CASE nCode OF
	16#000 : sText := '0: No error  ';
	16#001 : sText := '1: Internal error  ';
	16#002 : sText := '2: No Rtime  ';
	16#003 : sText := '3: Allocation locked memory error  ';
	16#004 : sText := '4: Insert mailbox error  ';
	16#005 : sText := '5: Wrong receive HMSG  ';
	16#006 : sText := '6: target port not found  ';
	16#007 : sText := '7: target machine not found  ';
	16#008 : sText := '8: Unknown command ID  ';
	16#009 : sText := '9: Bad task ID  ';
	16#00A : sText := '10: No IO  ';
	16#00B : sText := '11: Unknown AMS command  ';
	16#00C : sText := '12: Win 32 error  ';
	16#00D : sText := '13: Port not connected  ';
	16#00E : sText := '14: Invalid AMS length  ';
	16#00F : sText := '15: Invalid AMS Net ID  ';
	16#010 : sText := '16: Low Installation level  ';
	16#011 : sText := '17: No debug available  ';
	16#012 : sText := '18: Port disabled  ';
	16#013 : sText := '19: Port already connected  ';
	16#014 : sText := '20: AMS Sync Win32 error  ';
	16#015 : sText := '21: AMS Sync Timeout  ';
	16#016 : sText := '22: AMS Sync AMS error  ';
	16#017 : sText := '23: AMS Sync no index map  '; 
	16#018 : sText := '24: Invalid AMS port  ';
	16#019 : sText := '25: No memory  ';
	16#01A : sText := '26: TCP send error  ';
	16#01B : sText := '27: Host unreachable  ';
	16#1000 : sText := '4096: Intern: RTERR_INTERNAL : $R$N Internal fatal error in the TwinCAT real-time system.  ';
	16#1001 : sText := '4097: Intern: RTERR_BADTIMERPERIODS: $R$N Timer value not vaild.  ';
	16#1002 : sText := '4098: Intern: RTERR_INVALIDTASKPTR: $R$N Task pointer has the invalid value ZERO. ';
	16#1003 : sText := '4099: Intern: RTERR_INVALIDSTACKPTR: $R$N Task stack pointer has the invalid value ZERO. ';
	16#1004 : sText := '4100: Intern: RTERR_PRIOEXISTS: $R$N The demand task priority is already assigned.  ';
	16#1005 : sText := '4101: Intern: RTERR_NOMORETCB: $R$N No more free TCB (Task Control Block) available. Maximum number of TCBs is 64.  ';
	16#1006 : sText := '4102: Intern: RTERR_NOMORESEMAS: $R$N No more free semaphores available. Maximum number of semaphores is 64.  ';
	16#1007 : sText := '4103: Intern: RTERR_NOMOREQUEUES: $R$N No more free queue available. Maximum number of queue is 64.  ';
	16#1008 : sText := '4104: Intern: TwinCAT reserved.:  ';
	16#1009 : sText := '4105: Intern: TwinCAT reserved.:  '; 
	16#100a : sText := '4106: Intern: TwinCAT reserved.:  '; 
	16#100b : sText := '4107: Intern: TwinCAT reserved.:  '; 
	16#100C : sText := '4108: Intern: TwinCAT reserved.:  ';
	16#100D : sText := '4109: Intern: RTERR_EXTIRQALREADYDEF: $R$N An external synchronisation interrupt is already applied. ';
	16#100E : sText := '4110: Intern: RTERR_EXTIRQNOTDEF: $R$N No external synchronsiation interrupt applied. ';
	16#100F : sText := '4111: Intern: RTERR_EXTIRQINSTALLFAILED: $R$N The apply of the external synchronisation interrupt failed. ';
	16#1010 : sText := '4112: Intern: RTERR_IRQLNOTLESSOREQUAL: $R$N Call of a service function in the wrong context.  ';
	16#2000 : sText := ': ERR_IOERRS  ';
	16#274C : sText := '10060: A socket operation was attempted to an unreachable host  ';
	16#274D : sText := '10061: A connection attempt failed because the connected party did not properly respond after a period of time, $R$N or established connection failed because connected host has failed to respond.  ';
	16#2751 : sText := '10065: No connection could be made because the target machine actively refused it  ';
	16#2900 : sText := ': ERR_DPSLAVE (ERR_IOERRS+0x900)  ';
	16#2A00 : sText := ': ERR_CP5412A2 (ERR_IOERRS+0xA00)  '; 
	16#2B00 : sText := ': ERR_ASP (ERR_IOERRS+0xB00)  '; 
	16#2C00 : sText := ': ERR_CANSLAVE (ERR_IOERRS+0xC00)  '; 
	16#2D00 : sText := ': ERR_CIF30 (ERR_IOERRS+0xD00)  '; 
	16#2E00 : sText := ': ERR_IBSSLAVE (ERR_IOERRS+0xE00)  ';
	16#3000 : sText := ': ERR_SPSERRS  '; 
	16#4000 : sText := ': ERR_NCERRS  ';
	16#500 : sText := '1280: Intern: ROUTERERR_NOLOCKEDMEMORY: $R$N No locked memory can be allocated.  ';
	16#501 : sText := '1281: Intern: ROUTERERR_RESIZEMEMORY: $R$N The size of the  router memory could not be changed. ';
	16#502 : sText := '1282: Intern: ROUTERERR_MAILBOXFULL: $R$N The Mailbox of the AmsPort has reached the maximum number of possible entries. The current sent message was abolished.  ';
	16#503 : sText := '1283: Intern: ROUTERERR_DEBUGBOXFULL: $R$N The Mailbox of the Ams debugger port has reached the maximum number of possible entries. $R$N The sent message wil not be displayed in the debug monitor.  ';
	16#504 : sText := '1284: Intern: ROUTERERR_UNKNOWNPORTTYPE :  ';
	16#505 : sText := '1285: Intern: ROUTERERR_NOTINITIALIZED: $R$N Router is not (yet) initialised.  ';
	16#506 : sText := '1286: Intern: ROUTERERR_PORTALREADYINUSE : $R$N The desired port number is already assigned. ';
	16#507 : sText := '1287: Intern: ROUTERERR_NOTREGISTERED : $R$N Ams Port not registered  ';
	16#508 : sText := '1288: Intern: ROUTERERR_NOMOREQUEUES: $R$N The maximum number of Ams Ports reached.  ';
	16#509 : sText := '1289: Intern: ROUTERERR_INVALIDPORT :  '; 
	16#50A : sText := '1290: Intern: ROUTERERR_NOTACTIVATED : $R$N TwinCAT Router not (yet) active.  ';
	16#6000 : sText := ': ERR_PLCERRS  ';
	16#0700 : sText := '1792: error class <device error>  ';
	16#7000 : sText := ': ERR_STRKERRS  '; 
	16#0701 : sText := '1793: Service is not supported by server  ';
	16#0702 : sText := '1794: invalid index group  ';
	16#0703 : sText := '1795: invalid index offset  ';
	16#0704 : sText := '1796: reading/writing not permitted  ';
	16#0705 : sText := '1797 : parameter size not correct  ';
	16#0706 : sText := '1798: invalid parameter value(s)  ';
	16#0707 : sText := '1799: device is not in a ready state  ';
	16#708 : sText := '1800: device is busy  '; 
	16#709 : sText := '1801: invalid context (must be in Windows)  ';
	16#70A : sText := '1802: out of memory  '; 
	16#70B : sText := '1803: invalid parameter value(s)  '; 
	16#70C : sText := '1804: not found (files, ...)  ';
	16#70D : sText := '1805: syntax error in command or file  '; 
	16#70E : sText := '1806: objects do not match  '; 
	16#70F : sText := '1807: object already exists  '; 
	16#710 : sText := '1808: symbol not found  '; 
	16#711 : sText := '1809: symbol version invalid  '; 
	16#712 : sText := '1810: server is in invalid state  '; 
	16#713 : sText := '1811: AdsTransMode not supported  '; 
	16#714 : sText := '1812: Notification handle is invalid  '; 
	16#715 : sText := '1813: Notification client not registered  '; 
	16#716 : sText := '1814: no more notification handles  '; 
	16#717 : sText := '1815: size for watch too big  ';
	16#718 : sText := '1816: device not initialized  ';
	16#719 : sText := '1817: device has a timeout  '; 
	16#71A : sText := '1818: query interface failed  '; 
	16#71B : sText := '1819: wrong interface required  '; 
	16#71C : sText := '1820: class ID is invalid  '; 
	16#71D : sText := '1821: object ID is invalid  '; 
	16#71E : sText := '1822: request is pending  '; 
	16#71F : sText := '1823: request is aborted  '; 
	16#720 : sText := '1824: signal warning  '; 
	16#721 : sText := '1825: invalid array index  ';
	16#722 : sText := '1826: symbol not active -> release handle and try again  ';
	16#723 : sText := '1827: access denied  ';
	16#740 : sText := '1856: Error class <client error>  ';
	16#741 : sText := '1857: invalid parameter at service  ';
	16#742 : sText := '1858: polling list is empty  '; 
	16#743 : sText := '1859: var connection already in use  ';
	16#744 : sText := '1860: invoke ID in use  ';
	16#745 : sText := '1861: timeout elapsed  ';
	16#746 : sText := '1862: error in win32 subsystem  '; 
	16#748 : sText := '1864: ads port not opened  '; 
	16#750 : sText := '1872: internal error in ads sync  ';
	16#751 : sText := '1873: hash table overflow  ';
	16#752 : sText := '1874: key not found in hash  ';
	16#753 : sText := '1875: no more symbols in cache  '; 
	16#754 : sText := '1876: invalid response received   ';
	16#755 : sText := '1877: Sync port locked: ADS-Client tries to send a ADS msg but another thread is still waiting for an ADS-response. $R$N This error occurs only if no ADS-router is installed (please install royalty free TwinCAT-CP) $R$N or the router does not know the remote ADS device (define the remote ADS partner )  ';
	16#7800 : sText := ': ERR_PRJSPECIFIC  ';
	ELSE
		sText := 'No Text for this ErrorCode available';
END_CASE;

F_AdsError_Text := sText;

END_FUNCTION

// ---- POUs/Tc3 Objects/Conversions/BitOriented/F_ConvArrBitsToWord_1.TcPOU
FUNCTION F_ConvArrBitsToWord_1 : WORD
VAR_INPUT
	arrBits: ARRAY [0..15] OF BOOL;
END_VAR
VAR
END_VAR

F_ConvArrBitsToWord := 0;

END_FUNCTION

// ---- POUs/Tc3 Objects/Diagnostic/Terminal/FB_TerminalDiagnosis_1.TcPOU
FUNCTION_BLOCK FB_TerminalDiagnosis_1
VAR_INPUT
	stTerminalState				:ST_TerminalState;
END_VAR
VAR_OUTPUT
	bTerminalOK					:BOOL;
	sTerminalStatus				:STRING;
END_VAR
VAR

	sStateStatusAll				:STRING(255);
	sState						:STRING;
	sWorkingState				:STRING;

END_VAR

(*This Function returns the State of the Device. Either one of the States INIT, PREOP, OP, BOOTSTRAP or SAFE-OP is returned. stState is given the Value of the Function. *)
sState:= FUN_StateReturn(state:= stTerminalState.unInfoState);

(*All other Errors that can occur concerning the State of the Device*)
(*Because theoratically all the other errors could occur all together, CONCAT is done to show them all in one view box.*)
IF stTerminalState.unInfoState.4
THEN
	sStateStatusAll:= 'Slave signals error. ';
ELSE
	sStateStatusAll:= '';
END_IF

IF stTerminalState.unInfoState.5
THEN
	sStateStatusAll:= CONCAT( sStateStatusAll, 'Invalid vendorID. ');
ELSE
	sStateStatusAll:= CONCAT( sStateStatusAll, '');
END_IF

IF stTerminalState.unInfoState.6
THEN
	sStateStatusAll:= CONCAT( sStateStatusAll, 'Initialization error occurred. ');
ELSE
	sStateStatusAll:= CONCAT( sStateStatusAll, '');
END_IF

IF stTerminalState.unInfoState.7
THEN
	sStateStatusAll:= CONCAT( sStateStatusAll, 'Slave disabled. ');
ELSE
	sStateStatusAll:= CONCAT( sStateStatusAll, '');
END_IF

IF stTerminalState.unInfoState.8
THEN
	sStateStatusAll:= CONCAT( sStateStatusAll, 'Slave not present. ');
ELSE
	sStateStatusAll:= CONCAT( sStateStatusAll, '');
END_IF

IF stTerminalState.unInfoState.9
THEN
	sStateStatusAll:= CONCAT( sStateStatusAll, 'Slave signals link error. ');
ELSE
	sStateStatusAll:= CONCAT( sStateStatusAll, '');
END_IF

IF stTerminalState.unInfoState.10
THEN
	sStateStatusAll:= CONCAT( sStateStatusAll, 'Slave signals missing link. ');
ELSE
	sStateStatusAll:= CONCAT( sStateStatusAll, '');
END_IF

IF stTerminalState.unInfoState.11
THEN
	sStateStatusAll:= CONCAT( sStateStatusAll, 'Slave signals unexpected link. ');
ELSE
	sStateStatusAll:= CONCAT( sStateStatusAll, '');
END_IF

IF stTerminalState.unInfoState.12
THEN
	sStateStatusAll:= CONCAT( sStateStatusAll,  'Communication port A. ');
ELSE
	sStateStatusAll:= CONCAT( sStateStatusAll, '');
END_IF

IF stTerminalState.unInfoState.13
THEN
	sStateStatusAll:= CONCAT( sStateStatusAll, 'Communication port B. ');
ELSE
	sStateStatusAll:= CONCAT( sStateStatusAll, '');
END_IF

IF stTerminalState.unInfoState.14
THEN
	sStateStatusAll:= CONCAT( sStateStatusAll, 'Communication port C. ');
ELSE
	sStateStatusAll:= CONCAT( sStateStatusAll, '');
END_IF

IF stTerminalState.unInfoState.15
THEN
	sStateStatusAll:= CONCAT( sStateStatusAll,  'Communication port D. ');
ELSE
	sStateStatusAll:= CONCAT( sStateStatusAll, '');
END_IF

(*If none of the other errors occur, the text of the view box is 'None'.*)
IF sStateStatusAll= ''
THEN
	sStateStatusAll:= 'No error';
END_IF

(*The colour and text of the view box WcState is adjusted.*)
IF stTerminalState.bWcState = 0
THEN
	sWorkingState:= 'Working State OK ';
ELSE
	sWorkingState:= 'Working State NOT OK ';
END_IF

(*General Status Information*)
IF stTerminalState.bWcState= 0
     AND sStateStatusAll= 'No error'
THEN
	bTerminalOK:= TRUE;
	sTerminalStatus:= 'Terminal OK ';
ELSE
	bTerminalOK:= FALSE;
	sTerminalStatus:= 'Terminal Error ';
END_IF

END_FUNCTION_BLOCK

// ---- POUs/Tc3 Objects/Diagnostic/Terminal/FUN_StateReturn.TcPOU
FUNCTION FUN_StateReturn : STRING
VAR_INPUT
	state: UINT;
END_VAR
VAR
END_VAR

(*This Function returns the State of the Device. Either one of the States INIT, PREOP, OP, BOOTSTRAP or SAFE-OP is returned.
FB_Diagnosis.stState is given the Value of this Function. *)

IF state.0 AND NOT state.1 THEN
	FUN_StateReturn:= 'Slave in INIT state';
END_IF
IF state.1 AND NOT state.0 THEN
	FUN_StateReturn:= 'Slave in PREOP state';
END_IF
IF state.0 AND state.1 THEN
	FUN_StateReturn:= 'Slave in BOOTSTRAP state';
END_IF
IF state.2 THEN
	FUN_StateReturn:= 'Slave in SAFEOP state';
END_IF
IF state.3 THEN
	FUN_StateReturn:= 'Slave in OP state';
END_IF

END_FUNCTION

// ---- POUs/Tc3 Objects/Diagnostic/Terminal/FB_ToggleBit_1.TcPOU
FUNCTION_BLOCK FB_ToggleBit_1
VAR_INPUT
(*+++++ TxPDO Toggle +++++*)
	bToggle: BOOL;
END_VAR
VAR_OUTPUT
END_VAR
VAR
(*+++++ Toggle Bit Bridge +++++*)
	rtToggle: R_TRIG;
	ftToggle: F_TRIG;
	rCounter: REAL;
	rLastCounter: REAL;
(*+++++ Evaluation of Toggle Bits +++++*)
	tonTimer: TON;
	rToggleBitCounter: REAL;
	rUpdateTime: REAL;
END_VAR

(*This function block evaluates the Toggle Bit of the device.
Within a period of 10 seconds, is is checked how often the Toggle Bit changes it's value. *)

rtToggle(CLK:= bToggle);
ftToggle(CLK:= bToggle);

tonTimer.IN:= TRUE;
tonTimer.PT:= t#10000ms;

IF NOT tonTimer.Q THEN
	IF rtToggle.Q THEN
		rCounter:= rCounter+1;
	END_IF
	IF ftToggle.Q THEN
		rCounter:= rCounter+1;
	END_IF

	rToggleBitCounter:= rCounter;
ELSE
	rLastCounter:= rCounter;
	rUpdateTime:= SEL(rLastCounter = 0, 1 / (rLastCounter/10), 0); 		(*Update Time is calculated*)
	rCounter:= 0;
	tonTimer.IN:= FALSE;
END_IF

tonTimer();

END_FUNCTION_BLOCK

// ---- POUs/Tc3 Objects/Engineering/Buffer/FB_FiFo_1.TcPOU
FUNCTION_BLOCK FB_FiFo_1
(*
FiFo buffer of strings.

Constructor: 		Patryk Panylo
Company:		E. Riexinger GmbH
Date:			14.05.2013
Version:			1.00

Date:			Revision:		Who:				Comment
dd.mm.yyyy		x.xx			Initials			comment

*)
VAR_INPUT
	bAdd				:BOOL;
	bClear				:BOOL;
	sItem				:STRING;
END_VAR
VAR_OUTPUT

END_VAR
VAR_IN_OUT
	arsBuffer				:ARRAY[0..unSize] OF STRING;			(* Circular buffer *)
END_VAR
VAR
	bNoBufferEmpty		:BOOL;									(* Buffer empty *)
	nIdx					:INT;

	rtAdd				:R_TRIG;
	rtClear				:R_TRIG;
END_VAR
VAR CONSTANT
	unSize				:UINT := 100;								(* Buffer size *)
END_VAR

(* Add date to buffor *)
rtAdd(CLK := bAdd);

IF rtAdd.Q
THEN
	FOR nIdx := unSize - 1 TO 0 BY -1
	DO
		arsBuffer[nIdx + 1] := arsBuffer[nIdx];
	END_FOR

	arsBuffer[0] := sItem;

	RETURN;
END_IF

(* Clear buffor *)
rtClear(CLK := bClear);

IF rtClear.Q
THEN
	MEMSET(ADR(arsBuffer), 0, SIZEOF(arsBuffer));
	nIdx := 0;
END_IF

END_FUNCTION_BLOCK

// ---- POUs/Tc3 Objects/Engineering/External set value generator/FB_ExtSetpoint_1.TcPOU
FUNCTION_BLOCK FB_ExtSetpoint_1
(*

The function block used to move axis with an external set value.

Constructor: 		Patryk Panylo
Company:		E. Riexinger GmbH
Date:			01.04.2015
Version:			1.00

Date:			Revision:		Who:				Comment
dd.mm.yyyy		x.xx			Initials			comment

*)
VAR_INPUT
	(* Input variables / Eingang Variablen *)
	bEnable						:BOOL;						(* Function block enable *)
	bNoEStop					:BOOL;						(* No ermergency Stop / Keine Notaus *)
	
	byConfig					:BYTE;						(* Bit 0 - external trajectory,
															   Bit 1 - 
		
															*)
	bStart						:BOOL;						(* Execute start an external set value generator with rising edge *)
	bStop						:BOOL;						(* Execute stop an external set value generator with rising edge *)
	lrPosition					:LREAL;						(* Set position from an external set value generator *)
	lrPositionOffset			:LREAL;						(* Set offset of position *)
	ePositionType 				:E_PositionType ;			(* Position type - POSITIONTYPE_ABSOLUTE or POSITIONTYPE_RELATIVE *)
	bNotMoving					:BOOL;						(* Set not moving *)
	bNegativeDirection			:BOOL;						(* Negative direction *)
	bPositiveDirection			:BOOL;						(* Positive direction *)
	lrVelocity					:LREAL;						(* Set velocity from an external set point generator  > 0 *)
	lrAcceleration				:LREAL;						(* Set acceleration from an external set point generator > 0 *)					
END_VAR
VAR_OUTPUT
	(* Output variables / Ausgang Variablen *)
	bEnabled  				:BOOL;						(* Enabled shows the current state of the external set point generator *)
	bDone					:BOOL;						(* Command done *)
	bBusy					:BOOL;						(* Command busy *)
	bError					:BOOL;						(* Command error  *)
	udnErrorNo				:UDINT;						(* Error number *)
	sErrorMsg				:STRING; 					(* Error message *)
END_VAR
VAR_IN_OUT
	AxisDest				:AXIS_REF;					(* The AXIS_REF data type  is an interface between the PLC and the NC and contains axis information *)
END_VAR
VAR
	(* Instances / Instanzen *)
	fbMC_ExtSetPointGenEnable			:MC_ExtSetPointGenEnable;						(* Switch on external set value generator with the function. *)
	fbMC_ExtSetPointGenDisable			:MC_ExtSetPointGenDisable;						(* Switch off external set value generator with the function. *)

	rtStart								:R_TRIG;
	rtStop								:R_TRIG;
	bExtStart							:BOOL;
	bExtStop							:BOOL;
	
	(* Enumerator  *)
	etExtSetpoint						:ET_ExtSetpoint;								(* Current state *)

	(* General flags / Allgemeine Variablen *)
	eLastPositionType 					:E_PositionType;
	lrExtPosition						:LREAL;
	lrExtVelocity						:LREAL;
	lrExtAcceleration					:LREAL;
	dnExtDirection						:DINT;
	bImediateStop						:BOOL;
	bFirstTime							:BOOL;

END_VAR
VAR CONSTANT
	lrEPSILON				 :LREAL := 1E-6;
END_VAR

IF NOT bEnable
THEN
	bDone := bStart OR bStop;			(* Command done *)
	bBusy := bStart OR bStop;			(* Command busy *)
	bError := FALSE;					(* Command error  *)
	udnErrorNo := 0;					(* Error number *)
	sErrorMsg := ''; 					(* Error message *)

	bEnabled := bStart;
	
	bFirstTime := FALSE;
	RETURN;
END_IF

IF NOT bFirstTime
THEN
	bEnabled := FALSE;

	fbMC_ExtSetPointGenEnable(Execute := FALSE, Axis := AxisDest);						(* Reset FB and get Enabled status *)
	fbMC_ExtSetPointGenDisable(Execute := FALSE, Axis := AxisDest); 						(* Reset FB and get Enabled status *)

	etExtSetpoint := ET_ExtSetpoint_eWaitExecute;

	bFirstTime := TRUE;
END_IF

bImediateStop := AxisInErrorState(AxisDest.NcToPlc.AxisState);
IF bImediateStop
THEN
	(* Stop generator if axis is in error state *)
	lrExtVelocity := 0.0;
	lrExtAcceleration := 0.0;
	dnExtDirection := 0;
	bError := TRUE;													(* Command error  *)
	udnErrorNo :=  AxisDest.NcToPlc.ErrorCode;						(* Error number *)
	sErrorMsg := ''; 												(* Error message *)

	etExtSetpoint := ET_ExtSetpoint_eError;

ELSE
	(* Produce the dynamic data for the external setpoint generator interface *)
	lrExtVelocity := lrVelocity;
	lrExtAcceleration := lrAcceleration;
END_IF

lrExtPosition :=  lrPosition + lrPositionOffset;

(*IF bNotMoving
THEN
	dnExtDirection := 0;				(* Stand still *)
ELS*)IF bNegativeDirection
THEN
	dnExtDirection := -1;				(* Negative motion *)	
ELSIF bPositiveDirection
THEN
	dnExtDirection := 1;				(* Positive motion *)
ELSE
	dnExtDirection := 0;				(* Positive motion *)
END_IF

rtStart(CLK := AxisDest.Status.Operational);
bExtStart := (bStart OR rtStart.Q); // AND AxisDest.Status.Operational;
//rtStop(CLK := dnExtDirection = 0);
bExtStop := bStop OR rtStop.Q OR (NOT bNoEStop AND bNotMoving);

IF rtStop.Q
THEN
	etExtSetpoint := ET_ExtSetpoint_eWaitExecute;
END_IF

CASE etExtSetpoint
OF
	ET_ExtSetpoint_eWaitExecute:
		IF bExtStop
		THEN
			fbMC_ExtSetPointGenEnable(Execute := FALSE, Axis := AxisDest);						(* Reset FB and get Enabled status *)
			fbMC_ExtSetPointGenDisable(Execute := FALSE, Axis := AxisDest); 					(* Reset FB and get Enabled status *)

			bDone := FALSE;						(* Command done *)
			bBusy := TRUE;						(* Command busy *)
			bError := FALSE;						(* Command error  *)
			udnErrorNo := 0;						(* Error number *)
			sErrorMsg := ''; 						(* Error message *)

			etExtSetpoint := ET_ExtSetpoint_eDisableExtSetPointGenerator;

		ELSIF bExtStart
		THEN
			fbMC_ExtSetPointGenEnable(Execute := TRUE, Axis := AxisDest);						(* Reset FB and get Enabled status *)
			fbMC_ExtSetPointGenDisable(Execute := FALSE, Axis := AxisDest); 					(* Reset FB and get Enabled status *)

			bDone := FALSE;						(* Command done *)
			bBusy := TRUE;						(* Command busy *)
			bError := FALSE;						(* Command error  *)
			udnErrorNo := 0;						(* Error number *)
			sErrorMsg := ''; 						(* Error message *)

			etExtSetpoint := ET_ExtSetpoint_eEnableExtSetPointGenerator;

			(* Check for errors *)
			(* lrExtVelocity < lrEPSILON
			THEN
				udnErrorNo := 1;						(* Error number *)

				etMoveExtState := ET_MoveExtState_eError;
			END_IF
			IF lrExtAcceleration < lrEPSILON
			THEN
				udnErrorNo := 2;						(* Error number *)

				etMoveExtState := ET_MoveExtState_eError;
			END_IF*)
		END_IF

	ET_ExtSetpoint_eEnableExtSetPointGenerator:
		IF fbMC_ExtSetPointGenEnable.Enabled
		    AND NOT fbMC_ExtSetPointGenEnable.Execute
		    AND (ePositionType = eLastPositionType)
		THEN
			(* Send enable command to set the new target position but do not wait until the command has finished *)
			fbMC_ExtSetPointGenEnable.Execute := TRUE ;
			fbMC_ExtSetPointGenEnable.PositionType := ePositionType;

			etExtSetpoint := ET_ExtSetpoint_eDone;

		ELSE
			(* Enable the set point generator *)
			fbMC_ExtSetPointGenEnable.Execute := TRUE ;
			fbMC_ExtSetPointGenEnable.PositionType := ePositionType;

			IF fbMC_ExtSetPointGenEnable.Error
			     AND NOT fbMC_ExtSetPointGenEnable.Busy
			THEN
				udnErrorNo := fbMC_ExtSetPointGenEnable.ErrorID;						(* Error number *)
				
				fbMC_ExtSetPointGenEnable.Execute := FALSE ;
						
				etExtSetpoint := ET_ExtSetpoint_eError;

			ELSIF fbMC_ExtSetPointGenEnable.Done
			      AND NOT fbMC_ExtSetPointGenEnable.Busy
			THEN
				fbMC_ExtSetPointGenEnable.Execute := FALSE ;
				
				eLastPositionType := ePositionType;

				etExtSetpoint := ET_ExtSetpoint_eDone;
			END_IF

		END_IF

	ET_ExtSetpoint_eDisableExtSetPointGenerator:
		(* Call the disable external set point generator function block *)
		fbMC_ExtSetPointGenDisable(Execute := TRUE, Axis := AxisDest);
		
		IF fbMC_ExtSetPointGenDisable.Error
		     AND NOT fbMC_ExtSetPointGenEnable.Busy
		THEN
			udnErrorNo := fbMC_ExtSetPointGenDisable.ErrorID;										(* Error number *)
			
			fbMC_ExtSetPointGenDisable(Execute := FALSE, Axis:=AxisDest);
		
			etExtSetpoint := ET_ExtSetpoint_eError;
		
		ELSIF fbMC_ExtSetPointGenDisable.Done
		      AND NOT fbMC_ExtSetPointGenEnable.Busy
		THEN
			fbMC_ExtSetPointGenDisable(Execute := FALSE, Axis:=AxisDest);
			
			etExtSetpoint := ET_ExtSetpoint_eDone;
		END_IF

	ET_ExtSetpoint_eError:
		bBusy := FALSE;						(* Command busy *)
		bError := TRUE;						(* Command error  *)

		etExtSetpoint := ET_ExtSetpoint_eNoExecute;

	ET_ExtSetpoint_eDone:
		bDone := TRUE;						(* Command done *)
		bBusy := FALSE;						(* Command busy *)

		etExtSetpoint := ET_ExtSetpoint_eNoExecute;

	ET_ExtSetpoint_eNoExecute:
		IF NOT bExtStart
		   AND NOT bExtStop
		THEN
			(* Reset outputs *)
			bDone := FALSE;						(* Command done *)
			bBusy := FALSE;						(* Command busy *)
			bError := FALSE;						(* Command error  *)

			etExtSetpoint := ET_ExtSetpoint_eWaitExecute;
		END_IF
END_CASE

bError := fbMC_ExtSetPointGenEnable.Error							(* Command error  *)
		  OR fbMC_ExtSetPointGenEnable.Error;

(* The function is used to feed set values from an external set point generator into an axis. *)
MC_ExtSetPointGenFeed(
	Position := lrExtPosition,
	Velocity := lrExtVelocity,
	Acceleration := lrExtAcceleration,
	Direction := dnExtDirection,
	Axis := AxisDest
);

(* Call the enable external set point generator function block *)
fbMC_ExtSetPointGenEnable(
	Position := lrPosition,
	Enabled => bEnabled,
	Axis := AxisDest
 );

END_FUNCTION_BLOCK

// ---- POUs/Tc3 Objects/Engineering/Filter/FB_PT1_1.TcPOU
FUNCTION_BLOCK FB_PT1_1
(*

Function block low-pass filter (PT1)  for damping of fast alternating input-values.
K(s) = k/1+sT1  -> h(t) = k(1 - e^(-t/T1))

The Discrete-Time Integrator using Euler method: 
y(n+1) = 1/T1 * dt * (kp * xn - yn) + yn => kp * xn * dt / T1+ yn * (1 - dt / T1)

y(n+1) = kp * xn * Tcycle / T1+ yn * (1 - Tcycle / T1)
T1 = 0 =>  y(n+1) = kp * xn

Sample Time
Constructor: 		Patryk Panylo
Company:		E. Riexinger GmbH
Date:			20.03.2014
Version:			1.00

Date:			Revision:		Who:				Comment
dd.mm.yyyy		x.xx			Initials			comment

*)
VAR_INPUT
	(* Variables *)
	bEnable								:BOOL;						(* Enable FB *)
	lrInSignal								:LREAL;						(* Input value to the block *)
	lrKp									:LREAL := 1;					(* Proportional gain of integrator *)
	tT1									:TIME := t#200ms;				(* Time constant  of integrator *)
	tTaskCycle							:TIME := t#10ms;				(* Cycle time *)
END_VAR
VAR_OUTPUT
	(* Variables *)
	lrOutSignal							:LREAL;						(* Output value the block state *)
END_VAR
VAR
	(* Variables *)
	bFirstTime							:BOOL;
	lrTimeRatio							:LREAL;

	lrLastSignal							:LREAL;						(* Last signal *)
END_VAR

IF NOT bEnable
THEN
	lrOutSignal := 0.0;
	bFirstTime := FALSE;
	RETURN;
END_IF


IF NOT bFirstTime
     OR tT1= t#0ms
     OR tT1 < (tTaskCycle + tTaskCycle)
THEN
	lrOutSignal := lrKp * lrInSignal;

	bFirstTime := TRUE;
ELSE
	lrTimeRatio := TIME_TO_LREAL(tTaskCycle) / TIME_TO_LREAL(tT1);

	lrOutSignal := (lrKp * lrInSignal * lrTimeRatio) + (lrLastSignal * (1 -  lrTimeRatio));
END_IF

lrLastSignal := lrOutSignal;

END_FUNCTION_BLOCK

// ---- POUs/Tc3 Objects/Engineering/Filter/FB_ValueFilter_1.TcPOU
FUNCTION_BLOCK FB_ValueFilter_1
(*

Function block for filtering current input-value.

Sample Time
Constructor: 		Patryk Panylo
Company:		E. Riexinger GmbH
Date:			16.07.2014
Version:			1.00

Date:			Revision:		Who:				Comment
dd.mm.yyyy		x.xx			Initials			comment

*)
VAR_INPUT
	(* Enummerations *)

	(* Variables *)
	bEnable								:BOOL := TRUE;					(* Enable FB *)

	lrInSignal								:LREAL;							(* Input signal *)
	lrDeltaMax							:LREAL := 100;					(* Maximum difference between two input values *)

	(* References *)

	(* Interfaces *)

	(* Instances *)

END_VAR
VAR_OUTPUT
	(* Enummerations *)
	
	(* Variables *)
	lrOutSignal							:LREAL;							(* Output signal *)

	(* References *)

	(* Interfaces *)

	(* Instances *)
END_VAR
VAR
	(* Enummerations *)
	
	(* Variables *)
	bFirstTime							:BOOL;							(* First cycle *)

	lrCacheInSignal						:LREAL;							(* Copy of input signal *)
	dnOverLimitCounter					:DINT;							(* Counter of over limit *)

	lrLastSignal							:LREAL;							(* Last signal in time N *)
	lrSignalN_1							:LREAL;							(* Signal in time N - 1 *)
	lrSignalN_2							:LREAL;							(* Signal in time N - 2 *)
	lrSignalN_3							:LREAL;							(* Signal in time N - 3 *)

	(* References *)

	(* Interfaces *)

	(* Instances *)




END_VAR

IF NOT bEnable
THEN
	lrOutSignal := lrInSignal;

	bFirstTime := FALSE;
	RETURN;
END_IF

IF NOT bFirstTime
THEN
	lrSignalN_3 := lrInSignal;
	lrSignalN_2 := lrInSignal;
	lrSignalN_1 := lrInSignal;
	lrLastSignal := lrInSignal;

	bFirstTime := TRUE;
END_IF

lrSignalN_3 := lrSignalN_2;
lrSignalN_2 := lrSignalN_1;
lrSignalN_1 := lrLastSignal;

lrCacheInSignal := lrInSignal;

IF ABS( lrCacheInSignal - lrSignalN_1 ) <= lrDeltaMax
THEN
	lrLastSignal := lrCacheInSignal;
	dnOverLimitCounter := 0;

ELSE
	dnOverLimitCounter := dnOverLimitCounter + 1;

	IF dnOverLimitCounter <= 3
	THEN
		lrLastSignal	:= lrSignalN_1 + ((lrSignalN_1 - lrSignalN_2) + (lrSignalN_2 - lrSignalN_3)) / 2.0;

	ELSIF dnOverLimitCounter = 4
	THEN
		lrLastSignal := lrSignalN_1 + (lrCacheInSignal - lrSignalN_1) / 2.0;

	ELSE
		lrLastSignal := lrCacheInSignal;
	END_IF

END_IF

lrOutSignal := lrLastSignal;

END_FUNCTION_BLOCK

// ---- POUs/Tc3 Objects/Engineering/Position offset/F_PosOffset_1.TcPOU
FUNCTION F_PosOffset_1 : LREAL
(*

The function used to calculate position offset in range.

Constructor: 		Patryk Panylo
Company:		E. Riexinger GmbH
Date:			01.04.2015
Version:			1.00

Date:			Revision:		Who:				Comment
dd.mm.yyyy		x.xx			Initials			comment

*)
VAR_INPUT
	(* Input variables / Eingang Variablen *)
	bEnable							:BOOL;						(* Function enable *)
	lrCurrentPosHorizontal				:LREAL;						(* Current position of horizontal axis *)
	lrPosOffsetHorizontal				:LREAL;						(* Position offset of horizontal axis*)
	lrPosOffsetVertical					:LREAL;						(* Position offset of horizontal axis*)
	lrRangeOffset						:LREAL;						(* Range offset *)
END_VAR
VAR
	(* Variables *)

END_VAR

IF NOT bEnable
THEN
	F_PosOffset := 0.0;

	RETURN;
END_IF

IF  lrRangeOffset > 0.0
     AND lrCurrentPosHorizontal >= lrPosOffsetHorizontal - ABS(lrRangeOffset * 0.5)
     AND lrCurrentPosHorizontal <= lrPosOffsetHorizontal + ABS(lrRangeOffset * 0.5)
THEN
	F_PosOffset := lrPosOffsetVertical;
ELSE
	F_PosOffset := 0.0;
END_IF

END_FUNCTION

// ---- POUs/Tc3 Objects/Engineering/Position/F_ModuloDistance_1.TcPOU
FUNCTION F_ModuloDistance_1 : DINT
(*
Function for calculate modulo distance.

Constructor: 	Patryk Panylo
Company:		E. Riexinger GmbH
Date:			20.01.2014
Version:		1.00

Date:			Revision:		Who:				Comment
dd.mm.yyyy		x.xx			Initials			comment

*)

VAR_INPUT
	dwCurrentValue			:DWORD;
	dwOldValue				:DWORD;
	dwModuloValue			:DWORD;
END_VAR
VAR
	dwPosDistance			:DWORD;

END_VAR


F_ModuloDistance := DWORD_TO_DINT(dwCurrentValue - dwOldValue);

IF dwModuloValue <> 0
THEN
	dwPosDistance := F_ModDW(dwCurrentValue - dwOldValue, dwModuloValue);
	
	F_ModuloDistance := DWORD_TO_DINT(dwPosDistance);
	
	IF dwPosDistance > (dwModuloValue / 2) 
	THEN
		F_ModuloDistance := -DWORD_TO_DINT(dwModuloValue - dwPosDistance);
	END_IF
	
END_IF

END_FUNCTION

// ---- POUs/Tc3 Objects/ExternalHardware/Gefran/FB_GFX4IRCtrlZone_1.TcPOU
FUNCTION_BLOCK FB_GFX4IRCtrlZone_1
(*

The function block used to control Gerfan GFX4IR zone.

Constructor: 		Patryk Panylo
Company:		E. Riexinger GmbH
Date:			12.07.2016
Version:			1.00

Date:			Revision:		Who:				Comment
dd.mm.yyyy		x.xx			Initials			comment

*)
VAR_INPUT
	(* Input variables / Eingang Variablen *)
	bEnable							:BOOL;						(* Function block enable *)
	bReset							:BOOL;						(* Controller reset *)
	bPowerEnabled					:BOOL;						(* Power enabled *)
	bHandStart						:BOOL;						(* Execute start an external trajectory with rising edge *)
	bHandStop						:BOOL;						(* Execute stop an external trajectory with rising edge *)
	bAutoStart						:BOOL;						(* Execute start an external trajectory with rising edge *)
	bAutoStop						:BOOL;						(* Execute stop an external trajectory with rising edge *)
	bExeStop						:BOOL;						(* Execute stop *)
	bStartRelease					:BOOL;						(* Start release *)
	bCtrlInterrupt					:BOOL;						(* Control interrupt *)
	lrSetpoint						:LREAL;						(* Setpoint 0 - 100 *)
	bCtrlManAuto					:BOOL;						(* Auto := TRUE, Man := FALSE *)
	bEnAutoCtrlOff					:BOOL := TRUE;				(* Auto off enable*)
	tControllerOff					:TIME := T#90S;				(* Time to switch controller off *)
	tControllerOn					:TIME := T#90S;				(* Time to switch controller on *)
END_VAR
VAR_OUTPUT
	(* Output variables / Ausgang Variablen *)
	lrCurrentValue					:LREAL;						(* Current value *)
	bPowerEnable		 			:BOOL;						(* Power enable *)
	bSwitchOn		 				:BOOL;						(* Zone switch on *)
	bEnabled  						:BOOL;						(* Zone enabled *)
	bDamaged						:BOOL;						(* Zone damaged *)
	bDone							:BOOL;						(* Command done *)
	bBusy							:BOOL;						(* Command busy *)
	bError							:BOOL;						(* Command error  *)
	udnErrorNo						:UDINT;						(* Error number *)
	sErrorMsg						:STRING; 					(* Error message *)
END_VAR
VAR_IN_OUT
	(* Input Output variables / Ausgang Variablen *)
	CtrlGFX4IRTOPLC					:ST_GFX4IRTOPLC;			(* The ST_GFX4IRTOPLC data type  is an interface between the PLC and the GFX4IR and contains controller information *)
	CtrlPLCTOGFX4IR					:ST_PLCTOGFX4IR;			(* The ST_PLCTOGFX4IR data type  is an interface between the PLC and the GFX4IR and contains controller information *)
END_VAR
VAR
	(* Enummerations *)
	etGFX4IRStates					:ET_GFX4IR := ET_GFX4IRState_eWaitExecute;			(* Current state *)

	(* Variables *)
	bStop 							:BOOL;
	nWatchdog						:INT;
	bControllerOn					:BOOL;

	bFirstTime						:BOOL;

	(* References *)

	(* Interfaces *)

	(* Instances *)
	tofCtrlOn						:TOF;
	tonSwitchOn						:TON;
	tonDamaged						:TON;
	tonEnabled						:TON;			
	
	fbControllerOff					:FB_SignalHandlingDelay;
	fbControllerOn					:FB_SignalHandlingDelay;

	rtAutoStart						:R_TRIG;
	rtAutoStop						:R_TRIG;
	rtHandStart						:R_TRIG;
	rtHandStop						:R_TRIG;
	rtExeStop						:R_TRIG;
END_VAR
VAR CONSTANT
	tPowerOn						:TIME := T#500MS;
	tSwitchOn						:TIME := T#500MS;
	tEnabled						:TIME := T#2S500MS;
	tDamaged						:TIME := t#2s;
END_VAR


IF NOT bFirstTime
THEN
	IF bCtrlManAuto
	THEN
		CtrlPLCTOGFX4IR.wControllerStatus.4 := FALSE;			(* Auto *)
	ELSE
		CtrlPLCTOGFX4IR.wControllerStatus.4 := TRUE;			(* Manual *)
	END_IF

	bControllerOn := TRUE;

	bStop := TRUE;
	
	CtrlPLCTOGFX4IR.wControllerStatus.3 := TRUE;			(* Ctrl ON = FALSE, OFF = TRUE *)
	CtrlPLCTOGFX4IR.nLocalSetPoint := 0;
	CtrlPLCTOGFX4IR.nManualOutput := 0;

	nWatchdog := 0;
	bDone := FALSE;						(* Command done *)
	bBusy := FALSE;						(* Command busy *)
	bError := FALSE;						(* Command error  *)

	etGFX4IRStates := ET_GFX4IRState_eWaitExecute;

	bFirstTime := TRUE;
END_IF

tofCtrlOn(
	IN := NOT CtrlPLCTOGFX4IR.wControllerStatus.3,
	PT := tPowerOn
);

bPowerEnable := tofCtrlOn.Q
				AND NOT CtrlPLCTOGFX4IR.wControllerStatus.3			(* Ctrl ON = FALSE, OFF = TRUE *)
				AND NOT bCtrlInterrupt
     			AND NOT fbControllerOff.bOut
				AND NOT bStop;
tonSwitchOn(
	IN := bPowerEnable
		  AND bPowerEnabled,
	PT := tSwitchOn
);
bSwitchOn := tonSwitchOn.Q;

tonEnabled(
	IN := bSwitchOn
		  AND CtrlGFX4IRTOPLC.nOutputPower > 0
		  AND (LREAL_TO_INT(lrSetpoint  * 10) = CtrlGFX4IRTOPLC.nOutputPower),
		  (*AND CtrlGFX4IRTOPLC.wControllerStatus.5					(* Ctrl enabled  *)
			AND NOT CtrlGFX4IRTOPLC.wControllerStatus.0;			(* Alarm  *)*)
	PT:= tEnabled
);
bEnabled := tonEnabled.Q;

tonDamaged(
	IN := bSwitchOn
		  AND CtrlGFX4IRTOPLC.wControllerStatus.12,
	PT := tDamaged
);

bDamaged := tonDamaged.Q;
lrCurrentValue := CtrlGFX4IRTOPLC.nOutputPower * 0.1;

fbControllerOff(
	bEnable := TRUE,
	bIn := bEnAutoCtrlOff
		  AND bEnabled,
	tDelay := tControllerOff
);

fbControllerOn(
	bEnable := TRUE,
	bIn := NOT bEnabled					(* Ctrl disabled *)
		  AND NOT bControllerOn,
	tDelay := tControllerOn
);

(*
IF bHandStop
    OR bCtrlInterrupt
THEN
	CtrlPLCTOGFX4IR.wControllerStatus.3 := TRUE;			(* Ctrl ON = FALSE, OFF = TRUE *)
	CtrlPLCTOGFX4IR.nLocalSetPoint := 0;
	CtrlPLCTOGFX4IR.nManualOutput := 0;
ELSIF bHandStart
THEN
	CtrlPLCTOGFX4IR.wControllerStatus.3 := FALSE;			(* Ctrl ON = FALSE, OFF = TRUE *)
	CtrlPLCTOGFX4IR.nManualOutput := LREAL_TO_INT(lrSetpoint  * 10);
END_IF

RETURN;
*)

IF bCtrlInterrupt
     OR fbControllerOff.bOut
THEN
	bControllerOn := FALSE;

	bStop := TRUE;
	
	CtrlPLCTOGFX4IR.wControllerStatus.3 := TRUE;			(* Ctrl ON = FALSE, OFF = TRUE *)
	CtrlPLCTOGFX4IR.nLocalSetPoint := 0;
	CtrlPLCTOGFX4IR.nManualOutput := 0;

	nWatchdog := 0;
	bDone := FALSE;						(* Command done *)
	bBusy := FALSE;						(* Command busy *)
	bError := FALSE;						(* Command error  *)

	etGFX4IRStates := ET_GFX4IRState_eWaitExecute;

ELSIF fbControllerOn.bOut
THEN
	bControllerOn := TRUE;
END_IF

IF bReset
     AND bError
THEN
	(* Reset outputs *)
	nWatchdog := 0;
	bDone := FALSE;						(* Command done *)
	bBusy := FALSE;						(* Command busy *)
	bError := FALSE;						(* Command error  *)

	etGFX4IRStates := ET_GFX4IRState_eWaitExecute;
ELSE
	(*IF bEnable
	     AND CtrlGFX4IRTOPLC.wControllerStatus.8					(* Ctrl error *)
	THEN
		bError := TRUE;									(* Command error  *)

		etGFX4IRStates := ET_GFX4IRState_eError;             		(* Next step *)
	END_IF*);
END_IF

rtHandStart(CLK := bHandStart);
rtHandStop(CLK := bHandStop);
rtAutoStart(CLK := bAutoStart AND bStartRelease AND bControllerOn);
rtAutoStop(CLK := bAutoStop);
rtExeStop(CLK := bExeStop);

IF rtExeStop.Q
	OR rtAutoStart.Q OR rtAutoStop.Q
THEN
	nWatchdog := 0;
	bDone := FALSE;						(* Command done *)
	bBusy := FALSE;						(* Command busy *)
	bError := FALSE;						(* Command error  *)

	bStop := TRUE;

	etGFX4IRStates := ET_GFX4IRState_eWaitExecute;	

ELSIF rtHandStart.Q OR rtHandStop.Q 
THEN
	nWatchdog := 0;
	bDone := FALSE;						(* Command done *)
	bBusy := FALSE;						(* Command busy *)
	bError := FALSE;						(* Command error  *)

	bStop := FALSE;

	etGFX4IRStates := ET_GFX4IRState_eWaitExecute;
END_IF

CASE etGFX4IRStates
OF
	ET_GFX4IRState_eWaitExecute:
		IF NOT bEnable
		THEN
			bDone := TRUE;						(* Command done *)
			bBusy := TRUE;						(* Command busy *)
			bError := FALSE;						(* Command error  *)
			bEnabled  := bAutoStart AND NOT bAutoStop; 				(* Controller enabled *)

			bStop := TRUE;
			
			CtrlPLCTOGFX4IR.wControllerStatus.3 := TRUE;			(* Ctrl ON = FALSE, OFF = TRUE *)
			CtrlPLCTOGFX4IR.nLocalSetPoint := 0;
			CtrlPLCTOGFX4IR.nManualOutput := 0;

			etGFX4IRStates := ET_GFX4IRState_eWaitExecute;

		ELSE
			IF rtExeStop.Q
			   OR bAutoStop
			   OR bHandStop
			THEN
				nWatchdog := 0;

				bDone := FALSE;						(* Command done *)
				bBusy := TRUE;						(* Command busy *)
				bError := FALSE;						(* Command error  *)
				udnErrorNo := 0;						(* Error number *)
				sErrorMsg := ''; 						(* Error message *)

				etGFX4IRStates := ET_GFX4IRState_eCtrlOff;

			ELSIF (rtAutoStart.Q
				   OR (rtHandStart.Q
					    AND bStartRelease
					    AND bControllerOn))
				   AND NOT bCtrlInterrupt
				   AND NOT fbControllerOff.bOut
			THEN
				nWatchdog := 0;
	
				bDone := FALSE;						(* Command done *)
				bBusy := TRUE;						(* Command busy *)
				bError := FALSE;						(* Command error  *)
				udnErrorNo := 0;						(* Error number *)
				sErrorMsg := ''; 						(* Error message *)

				etGFX4IRStates := ET_GFX4IRState_eCtrlOn;

			END_IF
		END_IF

	ET_GFX4IRState_eCtrlOn:
		nWatchdog := nWatchdog + 1;
		IF nWatchdog > 25000
		THEN
			etGFX4IRStates := ET_GFX4IRState_eError;            		 (* Next step *)
		END_IF;

		bStop := FALSE;
		
		CtrlPLCTOGFX4IR.wControllerStatus.3 := FALSE;			(* Ctrl ON = FALSE, OFF = TRUE *)

		IF bCtrlManAuto
		THEN
			CtrlPLCTOGFX4IR.nLocalSetPoint := LREAL_TO_INT(lrSetpoint * 10);
		ELSE
			CtrlPLCTOGFX4IR.nManualOutput := LREAL_TO_INT(lrSetpoint  * 10);
		END_IF
		
		IF bEnabled											(* Ctrl enabled *)
		THEN
			nWatchdog := 0;
			etGFX4IRStates := ET_GFX4IRState_eDone;
		END_IF

	ET_GFX4IRState_eCtrlOff:
		nWatchdog := nWatchdog + 1;
		IF nWatchdog > 1000
		THEN
			etGFX4IRStates := ET_GFX4IRState_eError;             		(* Next step *)
		END_IF;

		bStop := TRUE;
		
		CtrlPLCTOGFX4IR.wControllerStatus.3 := TRUE;			(* Ctrl ON = FALSE, OFF = TRUE *)
		CtrlPLCTOGFX4IR.nLocalSetPoint := 0;
		CtrlPLCTOGFX4IR.nManualOutput := 0;

		IF NOT bEnabled
		THEN
			nWatchdog := 0;
			etGFX4IRStates := ET_GFX4IRState_eDone;
		END_IF

	ET_GFX4IRState_eDone:
		nWatchdog := 0;
		bDone := TRUE;						(* Command done *)
		bBusy := FALSE;						(* Command busy *)

		etGFX4IRStates := ET_GFX4IRState_eNoExecute;

	ET_GFX4IRState_eError:
		nWatchdog := 0;
		bBusy := FALSE;						(* Command busy *)
		bError := TRUE;						(* Command error  *)

		bStop := TRUE;
		
		CtrlPLCTOGFX4IR.wControllerStatus.3 := TRUE;			(* Ctrl ON = FALSE, OFF = TRUE *)
		CtrlPLCTOGFX4IR.nLocalSetPoint := 0;
		CtrlPLCTOGFX4IR.nManualOutput := 0;

		etGFX4IRStates := ET_GFX4IRState_eNoExecute;

	ET_GFX4IRState_eNoExecute:
		IF NOT bHandStart
		   AND NOT bHandStop
		   AND NOT bAutoStart
		   AND NOT bAutoStop
		THEN
			(* Reset outputs *)
			nWatchdog := 0;
			bDone := FALSE;						(* Command done *)
			bBusy := FALSE;						(* Command busy *)
			bError := FALSE;						(* Command error  *)

			etGFX4IRStates := ET_GFX4IRState_eWaitExecute;
		END_IF
END_CASE

END_FUNCTION_BLOCK

// ---- POUs/Tc3 Objects/ExternalHardware/Gefran/FB_GFX4IRZones_1.TcPOU
FUNCTION_BLOCK FB_GFX4IRZones_1
(*

The function block used to control Gerfan GFX4IR Zones.

Constructor: 		Patryk Panylo
Company:		E. Riexinger GmbH
Date:			12.07.2016
Version:			1.00

Date:			Revision:		Who:				Comment
dd.mm.yyyy		x.xx			Initials			comment

*)
VAR_INPUT
	(* Input variables / Eingang Variablen *)
	bEnable							:BOOL;													(* Function block enable *)
	arbZoneEn						:ARRAY[1..GVL_GFX4IR.nZONES_MAX_NO] OF BOOL;			(* Zone enable *)
	bReset							:BOOL;													(* Reset *)
	bPowerEnabled					:BOOL;													(* Power enabled *)
	bTerminalOK						:BOOL;													(* Terminal Ok *)
	arbHandStart					:ARRAY[1..GVL_GFX4IR.nZONES_MAX_NO] OF BOOL;			(* Execute start GFX4IR controller with rising edge *)
	arbHandStop						:ARRAY[1..GVL_GFX4IR.nZONES_MAX_NO] OF BOOL;			(* Execute stop GFX4IR controller with rising edge *)
	bAutoStart						:BOOL;													(* Execute start GFX4IR controller with rising edge *)
	bAutoStop						:BOOL;													(* Execute stop GFX4IR controller with rising edge *)
	bExeStop						:BOOL;													(* Execute stop *)
	bStartRelease					:BOOL;													(* Start release *)
	bCtrlInterrupt					:BOOL;													(* Control interrupt *)
	arlrSetpoint					:ARRAY[1..GVL_GFX4IR.nZONES_MAX_NO] OF LREAL;			(* Setpoint 0 - 100 *)
	bCtrlManAuto					:BOOL;													(* Auto := TRUE, Man := FALSE *)
	bEnAutoCtrlOff					:BOOL := TRUE;											(* Auto controller off enable*)
	bEnOneByOneOn					:BOOL := FALSE;											(* One by one switch on *)
	tDelayZoneOn					:TIME := T#100MS;										(* Delay time of zone one by one to switch on *)
	tControllerOff					:TIME := T#90S;											(* Time to switch controller off *)
	tControllerOn					:TIME := T#90S;											(* Time to switch controller on *)
END_VAR
VAR_OUTPUT
	(* Output variables / Ausgang Variablen *)
	arlrCurrentValue				:ARRAY[1..GVL_GFX4IR.nZONES_MAX_NO] OF LREAL;			(* Current value *)
	bPowerEnable					:BOOL;						(* Power enable *)
	bSwitchOn		 				:BOOL;						(* Zones switch on *)
	bEnabled  						:BOOL;						(* Zone enabled *)
	bEnabledDelay					:BOOL;						(* Zone enabled delay *)
	byZoneDamaged					:BYTE;						(* Zone damaged *)
	bDone							:BOOL;						(* Command done *)
	bError							:BOOL;						(* Command error  *)
	udnErrorNo						:UDINT;						(* Error number *)
END_VAR
VAR_IN_OUT
	(* Input Output variables / Ausgang Variablen *)
	GFX4IR							:ST_GFX4IR_REF;				(* The ST_GFX4IR_REF data type  is an interface between the PLC and the GFX4IR and contains controller information *)
END_VAR
VAR
	(* Enummerations *)

	(* Variables *)
	nIdx							:INT;
	tEnabledDelay					:TIME := T#1S;					(* Enabled delay time *)
	arbZoneDamaged					:ARRAY[1..GVL_GFX4IR.nZONES_MAX_NO] OF BOOL;

	bFirstTime						:BOOL;

	(* References *)

	(* Interfaces *)

	(* Instances *)
	arfbGFX4IRCtrlZone				:ARRAY[1..GVL_GFX4IR.nZONES_MAX_NO] OF FB_GFX4IRCtrlZone;
	tonEnabledDelay					:TON;						(* Delay controller enabled status *)
	tonDelayZoneOn					:ARRAY[1..GVL_GFX4IR.nZONES_MAX_NO] OF TON;						(* Delay zone one by one to switch on *)

END_VAR


IF NOT bEnable
THEN
	bDone := FALSE;					(* Command done *)
	bError := FALSE;					(* Command error  *)

	FOR nIdx := 1 TO GVL_GFX4IR.nZONES_MAX_NO
	DO
		arfbGFX4IRCtrlZone[nIdx](
			bAutoStart := bAutoStart,
			bAutoStop := bAutoStop,
			bCtrlInterrupt := bCtrlInterrupt,
			CtrlGFX4IRTOPLC := GFX4IR.Gfx4IRToPlc[nIdx],
			CtrlPLCTOGFX4IR := GFX4IR.PlcToGfx4IR[nIdx],
			lrCurrentValue => arlrCurrentValue[nIdx]
		 );
	END_FOR

	bSwitchOn := FALSE;
	bEnabled := FALSE;
	bEnabledDelay := FALSE;

	bFirstTime := FALSE;
	RETURN;
END_IF

IF NOT bFirstTime
THEN
	bDone := FALSE;					(* Command done *)
	bError := FALSE;					(* Command error  *)

	bPowerEnable := FALSE;
	bSwitchOn := FALSE;
	bEnabled := FALSE;
	bEnabledDelay := FALSE;

	bFirstTime := TRUE;
END_IF

byZoneDamaged := 0;
bPowerEnable := FALSE;
bSwitchOn := FALSE;
bEnabled := TRUE;
bDone := TRUE;
bError := FALSE;

FOR nIdx := 1 TO GVL_GFX4IR.nZONES_MAX_NO
DO
	
	IF bAutoStart
	THEN
		IF bEnOneByOneOn
		     AND tDelayZoneOn > t#0ms
		     AND nIdx > 1
		     AND NOT arfbGFX4IRCtrlZone[nIdx].bEnabled
		THEN
			tonDelayZoneOn[nIdx](
				IN := arfbGFX4IRCtrlZone[nIdx - 1].bEnable,
				PT := tDelayZoneOn
			);
	
			IF tonDelayZoneOn[nIdx].Q
			THEN
				arfbGFX4IRCtrlZone[nIdx].bStartRelease := bStartRelease;
			ELSE
				arfbGFX4IRCtrlZone[nIdx].bStartRelease := FALSE;;
			END_IF
		ELSE
			tonDelayZoneOn[nIdx](IN := FALSE);
			arfbGFX4IRCtrlZone[nIdx].bStartRelease := bStartRelease;
		END_IF
	ELSE
		tonDelayZoneOn[nIdx](IN := FALSE);
		arfbGFX4IRCtrlZone[nIdx].bStartRelease := bStartRelease;
	END_IF
	

	//arfbGFX4IRCtrlZone[nIdx].bStartRelease := bStartRelease;

	arfbGFX4IRCtrlZone[nIdx](
		bEnable := arbZoneEn[nIdx],
		bReset := bReset,
		bPowerEnabled := bPowerEnabled,
		bHandStart := arbHandStart[nIdx],
		bHandStop := arbHandStop[nIdx],
		bAutoStart := bAutoStart,
		bAutoStop := bAutoStop,
		bExeStop := bExeStop,
		bCtrlInterrupt := NOT bTerminalOK
						  OR bCtrlInterrupt,
		lrSetpoint := arlrSetpoint[nIdx],
		bCtrlManAuto := bCtrlManAuto,
		bEnAutoCtrlOff := bEnAutoCtrlOff,
		tControllerOff := tControllerOff,
		tControllerOn := tControllerOn,
		CtrlGFX4IRTOPLC := GFX4IR.Gfx4IRToPlc[nIdx],
		CtrlPLCTOGFX4IR := GFX4IR.PlcToGfx4IR[nIdx],
		lrCurrentValue => arlrCurrentValue[nIdx],
		bDamaged => arbZoneDamaged[nIdx]
	 );

	bPowerEnable := bPowerEnable OR arfbGFX4IRCtrlZone[nIdx].bPowerEnable;
	bSwitchOn := bSwitchOn OR arfbGFX4IRCtrlZone[nIdx].bSwitchOn;
	bEnabled := bEnabled AND arfbGFX4IRCtrlZone[nIdx].bEnabled;
	bDone := bDone AND arfbGFX4IRCtrlZone[nIdx].bDone;
	bError := bError OR arfbGFX4IRCtrlZone[nIdx].bError;

END_FOR

IF arbZoneDamaged[1] = TRUE
THEN
	byZoneDamaged.0 := TRUE;
ELSIF arbZoneDamaged[2] = TRUE
THEN
	byZoneDamaged.1 := TRUE;
ELSIF arbZoneDamaged[3] = TRUE
THEN
	byZoneDamaged.2 := TRUE;
ELSIF arbZoneDamaged[4] = TRUE
THEN
	byZoneDamaged.3 := TRUE;
END_IF

tonEnabledDelay(
	IN := bEnabled,
	PT := tEnabledDelay,
	Q => bEnabledDelay
);

END_FUNCTION_BLOCK

// ---- POUs/Tc3 Objects/ExternalHardware/Gefran/FB_GFX4IR_REF_1.TcPOU
FUNCTION_BLOCK FB_GFX4IR_REF_1
VAR_INPUT
	stTerminalState		AT %I*:ST_TerminalState;
	Gfx4IRToPlc			AT %I*:ARRAY[1..4] OF ST_GFX4IRTOPLC;
END_VAR
VAR_OUTPUT
	PlcToGfx4IR			AT %Q*:ARRAY[1..4] OF ST_PLCTOGFX4IR;
END_VAR
VAR
END_VAR

;

END_FUNCTION_BLOCK

// ---- POUs/Tc3 Objects/ExternalHardware/Gefran/F_ChkAllZonesNotEnabled_1.TcPOU
FUNCTION F_ChkAllZonesNotEnabled_1 : BOOL
(*

The function used to detect if all controller are enabled.

Constructor: 		Patryk Panylo
Company:		E. Riexinger GmbH
Date:			23.04.2015
Version:			1.00

Date:			Revision:		Who:				Comment
dd.mm.yyyy		x.xx			Initials			comment

*)
VAR_INPUT
	(* Input variables / Eingang Variablen *)
	bEnable						:BOOL;						(* Signal FB enable *)
	GFX4IR1						:ST_GFX4IR_REF;				(* The ST_GFX4IRTOPLC data type  is an interface between the PLC and the GFX4IR and contains controller information *)
	GFX4IR2						:ST_GFX4IR_REF;				(* The ST_GFX4IRTOPLC data type  is an interface between the PLC and the GFX4IR and contains controller information *)
	GFX4IR3						:ST_GFX4IR_REF;				(* The ST_GFX4IRTOPLC data type  is an interface between the PLC and the GFX4IR and contains controller information *)
	GFX4IR4						:ST_GFX4IR_REF;				(* The ST_GFX4IRTOPLC data type  is an interface between the PLC and the GFX4IR and contains controller information *)
END_VAR
VAR
	(* Enummerations *)

	(* Variables *)

	(* References *)

	(* Interfaces *)

	(* Instances *)

END_VAR


IF NOT bEnable							(* Signal FB enable *)
THEN
	F_ChkAllZonesNotEnabled := FALSE;

	RETURN;
END_IF

F_ChkAllZonesNotEnabled := GFX4IR1.Gfx4IRToPlc[1].nProcessVariable = 0
						   AND GFX4IR1.Gfx4IRToPlc[2].nProcessVariable = 0
						   AND GFX4IR1.Gfx4IRToPlc[3].nProcessVariable = 0
						   AND GFX4IR1.Gfx4IRToPlc[4].nProcessVariable = 0
						   AND GFX4IR2.Gfx4IRToPlc[1].nProcessVariable = 0
						   AND GFX4IR2.Gfx4IRToPlc[2].nProcessVariable = 0
						   AND GFX4IR2.Gfx4IRToPlc[3].nProcessVariable = 0
						   AND GFX4IR2.Gfx4IRToPlc[4].nProcessVariable = 0
						   AND GFX4IR3.Gfx4IRToPlc[1].nProcessVariable = 0
						   AND GFX4IR3.Gfx4IRToPlc[2].nProcessVariable = 0
						   AND GFX4IR3.Gfx4IRToPlc[3].nProcessVariable = 0
						   AND GFX4IR3.Gfx4IRToPlc[4].nProcessVariable = 0
						   AND GFX4IR4.Gfx4IRToPlc[1].nProcessVariable = 0
						   AND GFX4IR4.Gfx4IRToPlc[2].nProcessVariable = 0
						   AND GFX4IR4.Gfx4IRToPlc[3].nProcessVariable = 0
						   AND GFX4IR4.Gfx4IRToPlc[4].nProcessVariable = 0;

END_FUNCTION

// ---- POUs/Tc3 Objects/ExternalHardware/KUKA/FB_KUKA_Enable_1.TcPOU
FUNCTION_BLOCK FB_KUKA_Enable_1
(*

The function block used to move enable for an kuka

Constructor: 		Patryk Panylo
Company:		E. Riexinger GmbH
Date:			18.11.2016
Version:			1.00

Date:			Revision:		Who:				Comment

*)
VAR_INPUT
	(* Input variables / Eingang Variablen *)
	bEnable						:BOOL;			(* Signal FB enable *)
	bAutoHand					:BOOL;			(* Auto := TRUE, Hand := FALSE *)
	bNoEStop					:BOOL;			(* No ermergency Stop / Keine Notaus *)
	bMoveOn					:BOOL;			(* Enable the move enable *)
END_VAR
VAR_OUTPUT
	(* Output variables / Ausgang Variablen *)
	bMoveEnabled				:BOOL;			(* MoveEnabled = TRUE indicates that the kuka  drivers is ready for operation. *)
	bError						:BOOL;			(* Error *)
	udnErrorNo					:UDINT;			(* Error number *)
	sErrorMsg					:STRING; 		(* Error message *)
END_VAR
VAR_IN_OUT
	(* Input Output variables / Ausgang Variablen *)
	Kuka							:ST_KUKA_REF;
END_VAR
VAR
	(* Enummerations *)

	(* Variables *)
	tMoveEnabledDelay 					:TIME := t#300ms;

	(* References *)

	(* Interfaces *)

	(* Instances *)
	tonMoveEnabledDelay					:TON;
END_VAR


IF NOT bEnable
THEN
	Kuka.PlcToKuka.bMoveEnable := FALSE;                   		 (* Disable *)
	tonMoveEnabledDelay(IN := FALSE,
				    		 PT := tMoveEnabledDelay);
ELSE

	IF NOT bNoEStop
	THEN
		Kuka.PlcToKuka.bMoveEnable := FALSE;                   		 (* Disable *)

	ELSE
		IF bAutoHand			(* Auto *)
		THEN
			IF (bMoveOn
			      OR (NOT bMoveOn
				     AND Kuka.KukaToPlc.bInWorkArea))
			     AND Kuka.KukaToPlc.bIOActConf
			     AND Kuka.KukaToPlc.bExt
			THEN
				Kuka.PlcToKuka.bMoveEnable := TRUE;                   		 (* Enable *)
			ELSE
				Kuka.PlcToKuka.bMoveEnable := FALSE;                   		 (* Enable *)
			END_IF
		ELSE				(* Manual *)
			IF Kuka.KukaToPlc.bT1
			     OR Kuka.KukaToPlc.bT2
			     OR Kuka.KukaToPlc.bAut
			THEN
				Kuka.PlcToKuka.bMoveEnable := TRUE;                   		 (* Enable *)
			ELSE
				Kuka.PlcToKuka.bMoveEnable := FALSE;                   		 (* Enable *)
			END_IF
		END_IF
	END_IF;

END_IF;

tonMoveEnabledDelay(IN := Kuka.PlcToKuka.bMoveEnable,				(* Move enabled *)
			   		PT := tMoveEnabledDelay);
bMoveEnabled := tonMoveEnabledDelay.Q;

END_FUNCTION_BLOCK

// ---- POUs/Tc3 Objects/ExternalHardware/KUKA/FB_KUKA_Power_1.TcPOU
FUNCTION_BLOCK FB_KUKA_Power_1
(*

The function block used to enable drives for an kuka

Constructor: 		Patryk Panylo
Company:		E. Riexinger GmbH
Date:			18.11.2016
Version:			1.00

Date:			Revision:		Who:				Comment

*)
VAR_INPUT
	(* Input variables / Eingang Variablen *)
	bEnable						:BOOL;			(* Signal FB enable *)
	bNoEStop					:BOOL;			(* No ermergency Stop / Keine Notaus *)
	bDrivesOn					:BOOL;			(* Enable the drives *)
	lrOverride					:LREAL;			(* Velocity override in % for all motion commands. (0 <= Override <= 100.0) *)
END_VAR
VAR_OUTPUT
	(* Output variables / Ausgang Variablen *)
	bStatus						:BOOL;			(* Status = TRUE indicates that the axis is ready for operation. *)
	bError						:BOOL;			(* Error *)
	udnErrorNo					:UDINT;			(* Error number *)
	sErrorMsg					:STRING; 		(* Error message *)
END_VAR
VAR_IN_OUT
	(* Input Output variables / Ausgang Variablen *)
	Kuka						:ST_KUKA_REF;
END_VAR
VAR
	(* Enummerations *)

	(* Variables *)
	tStatusDelay 					:TIME := t#300ms;

	(* References *)

	(* Interfaces *)

	(* Instances *)
	tonStatusDelay				:TON;
END_VAR


IF NOT bEnable
THEN
	Kuka.PlcToKuka.bDrivesOn := FALSE;                   		 (* Switch on *)
	Kuka.PlcToKuka.bDrivesOff := FALSE;                   		 (* Switch off *)
	tonStatusDelay(IN := FALSE,
				    PT := tStatusDelay);
ELSE

	IF NOT bNoEStop
	     OR NOT bDrivesOn
	THEN
		Kuka.PlcToKuka.bDrivesOn := FALSE;                   		 (* Switch on *)
		Kuka.PlcToKuka.bDrivesOff := FALSE;                   		 (* Switch off *)
	ELSE
		IF Kuka.KukaToPlc.bIOActConf
		     AND NOT Kuka.KukaToPlc.bPeriRdy
		THEN
			Kuka.PlcToKuka.bDrivesOn := TRUE;                   	(* Switch on *)
			Kuka.PlcToKuka.bDrivesOff := TRUE;                   		 (* Switch off *)
		ELSE
			Kuka.PlcToKuka.bDrivesOn := FALSE;                   	 (* Switch on *)
			Kuka.PlcToKuka.bDrivesOff := TRUE;                   		 (* Switch off *)
		END_IF
	END_IF;

END_IF;

Kuka.PlcToKuka.nOverride := LREAL_TO_INT(LIMIT(0,lrOverride,100));

tonStatusDelay(IN := Kuka.KukaToPlc.bPeriRdy,		(* Control enabled *)
			   PT := tStatusDelay);
bStatus := tonStatusDelay.Q;

END_FUNCTION_BLOCK

// ---- POUs/Tc3 Objects/ExternalHardware/KUKA/FB_KUKA_Prg_1.TcPOU
FUNCTION_BLOCK FB_KUKA_Prg_1
(*

The function block used to start kuka

Constructor: 		Patryk Panylo
Company:		E. Riexinger GmbH
Date:			18.11.2016
Version:			1.00

Date:			Revision:		Who:				Comment

*)
VAR_INPUT
	(* Input variables / Eingang Variablen *)
	bEnable						:BOOL;			(* Signal FB enable *)
	bReset						:BOOL;			(* Signal reset *)
	bAutoHome					:BOOL;			(* Auto := TRUE, Home := FALSE *)
	bStart						:BOOL;			(* Start program *)
	bStop						:BOOL;			(* Stop program *)
	nProgNo						:INT;			(* Program number *)
	tMaxRefTime					:TIME := t#60s;	(* Maximal referenc time *)
END_VAR
VAR_OUTPUT
	(* Output variables / Ausgang Variablen *)
	bRunning					:BOOL;						(* Program running *)
	bDone						:BOOL;						(* Program done *)
	bBusy						:BOOL;						(* Program busy *)
	bError						:BOOL;						(* Error *)
	udnErrorNo					:UDINT;
END_VAR
VAR_IN_OUT
	(* Input Output variables / Ausgang Variablen *)
	Kuka						:ST_KUKA_REF;
END_VAR
VAR
	(* Enummerations *)
	etKukaStart					:ET_KukaStart;

	(* Variables *)
	bFirstTime					:BOOL;

	nWatchdog					:INT;

	(* References *)

	(* Interfaces *)

	(* Instances *)
	rtStart						:R_TRIG;
	rtStop						:R_TRIG;
	rtReset						:R_TRIG;
	tonWatchdog					:TON;

END_VAR


IF NOT bEnable
THEN
	bDone := FALSE;					(* Program done *)
	bBusy := FALSE;                                  	(* Program not busy *)
	bError := FALSE;                                 	(* Program not error *)
	udnErrorNo := 0;                                 		(* Error number *)

	Kuka.PlcToKuka.bPgReset := FALSE;
	Kuka.PlcToKuka.bExtStart := FALSE;
	Kuka.PlcToKuka.bPgNoParity := FALSE;
	Kuka.PlcToKuka.bPgNoValid := FALSE;

	RETURN;
END_IF;

IF NOT bFirstTime
THEN
	tonWatchdog(IN := FALSE);

	Kuka.PlcToKuka.bPgReset := FALSE;
	Kuka.PlcToKuka.bExtStart := FALSE;
	Kuka.PlcToKuka.bPgNoParity := FALSE;
	Kuka.PlcToKuka.bPgNoValid := FALSE;

	etKukaStart := ET_KukaStart_eWaitExecute;              (* Next step *)

	bFirstTime := TRUE;
END_IF

rtReset(CLK := bReset);

IF rtReset.Q
     AND bError
THEN
	bError := FALSE;

	tonWatchdog(IN := FALSE);

	Kuka.PlcToKuka.bPgReset := FALSE;
	Kuka.PlcToKuka.bExtStart := FALSE;
	Kuka.PlcToKuka.bPgNoParity := FALSE;
	Kuka.PlcToKuka.bPgNoValid := FALSE;

	etKukaStart := ET_KukaStart_eWaitExecute;              (* Next step *)
END_IF

(* Wait for triger *)
rtStart(
	CLK := bStart
);

IF rtStart.Q
     AND Kuka.PlcToKuka.bDrivesOff
     AND Kuka.PlcToKuka.bMoveEnable
     AND Kuka.KukaToPlc.bUserSafe
     AND Kuka.KukaToPlc.bAlarmStop
     AND Kuka.KukaToPlc.bPeriRdy
     AND NOT Kuka.KukaToPlc.bProAct
     AND NOT Kuka.PlcToKuka.bDrivesOn
     AND NOT Kuka.KukaToPlc.bStopMess
THEN
	Kuka.PlcToKuka.bPgReset := FALSE;
	Kuka.PlcToKuka.bExtStart := FALSE;
	Kuka.PlcToKuka.bPgNoParity := FALSE;
	Kuka.PlcToKuka.bPgNoValid := FALSE;
	Kuka.PlcToKuka.nPgNo := 0;

	etKukaStart := ET_KukaStart_eWaitExecute;              (* Next step *)

END_IF

rtStop(
	CLK := bStop
		    OR NOT Kuka.PlcToKuka.bDrivesOff
     		    OR NOT Kuka.PlcToKuka.bMoveEnable
     		    OR NOT Kuka.KukaToPlc.bUserSafe
     		    OR NOT Kuka.KukaToPlc.bAlarmStop
     		    OR NOT Kuka.KukaToPlc.bPeriRdy
     		    OR Kuka.PlcToKuka.bDrivesOn
     		    OR Kuka.KukaToPlc.bStopMess
);

IF rtStop.Q
THEN
	Kuka.PlcToKuka.bPgReset := TRUE;
	Kuka.PlcToKuka.bExtStart := FALSE;
	Kuka.PlcToKuka.bPgNoParity := FALSE;
	Kuka.PlcToKuka.bPgNoValid := FALSE;
	Kuka.PlcToKuka.nPgNo := 0;

	etKukaStart := ET_KukaStart_eWaitExecute;              (* Next step *)

ELSIF NOT Kuka.KukaToPlc.bApplRun
THEN
	Kuka.PlcToKuka.bPgReset := FALSE;
END_IF

bRunning := Kuka.KukaToPlc.bApplRun
		      AND Kuka.KukaToPlc.bProAct;

(* Send command *)
CASE etKukaStart OF

	ET_KukaStart_eWaitExecute:
		bBusy := FALSE;                                     	(* Program not busy *)
		bError := FALSE;                         		(* Program not error *)
		udnErrorNo := 0;                         		(* Error number *)

		IF rtStart.Q
		     AND NOT bStop
		THEN
			nWatchdog := 0;
			bDone:= FALSE;                               		(* Program done *)
			bBusy := TRUE;                                  	(* Program busy *)

			tonWatchdog(IN := FALSE);

			Kuka.PlcToKuka.bExtStart := FALSE;
			Kuka.PlcToKuka.bPgNoParity := FALSE;
			Kuka.PlcToKuka.bPgNoValid := FALSE;
			Kuka.PlcToKuka.nPgNo := nProgNo;

			IF NOT bAutoHome
			     AND Kuka.KukaToPlc.bInHome
			THEN
				etKukaStart := ET_KukaStart_eDone;              (* Next step *)
			ELSE
				etKukaStart := ET_KukaStart_eExtStart;              (* Next step *)
			END_IF

		END_IF

	ET_KukaStart_eExtStart:
		(*nWatchdog := nWatchdog + 1;*)

		Kuka.PlcToKuka.bExtStart := TRUE;
		Kuka.PlcToKuka.bPgNoParity := FALSE;
		Kuka.PlcToKuka.bPgNoValid := FALSE;

		IF Kuka.KukaToPlc.bProAct
		     AND Kuka.KukaToPlc.bOnPath
		     AND NOT Kuka.KukaToPlc.bApplRun
		     AND NOT Kuka.KukaToPlc.bStopMess
		THEN
			nWatchdog := 0;

			(*Kuka.PlcToKuka.bExtStart := FALSE;
			Kuka.PlcToKuka.bPgNoParity := FALSE;
			Kuka.PlcToKuka.bPgNoValid := FALSE;*)

			etKukaStart := ET_KukaStart_eWfInHome;              (* Next step *)

		ELSIF Kuka.KukaToPlc.bStopMess
			    OR nWatchdog > 1000
		THEN
			Kuka.PlcToKuka.bExtStart := FALSE;
			Kuka.PlcToKuka.bPgNoParity := FALSE;
			Kuka.PlcToKuka.bPgNoValid := FALSE;
			
			udnErrorNo := 1;                     (* Error number *)
			
			etKukaStart := ET_KukaStart_eError;              (* Next step *)

		END_IF

	ET_KukaStart_eWfInHome:
		tonWatchdog(
			IN := Kuka.PlcToKuka.nOverride > 0,
			PT:= tMaxRefTime
		);

		IF tonWatchdog.Q
		THEN
			tonWatchdog(IN := FALSE);

			Kuka.PlcToKuka.bExtStart := FALSE;
			Kuka.PlcToKuka.bPgNoParity := FALSE;
			Kuka.PlcToKuka.bPgNoValid := FALSE;

			udnErrorNo := 2;

			etKukaStart := ET_KukaStart_eError;             (* Next step *)

		ELSIF (NOT bAutoHome
			    OR (bAutoHome
				    AND (Kuka.KukaToPlc.bInHome
		     			       OR Kuka.KukaToPlc.arbInHome[1])))
			    AND Kuka.KukaToPlc.bProAct
		    	    AND Kuka.KukaToPlc.bOnPath
			    AND NOT Kuka.KukaToPlc.bApplRun
		     	    AND NOT Kuka.KukaToPlc.bStopMess
		THEN
			tonWatchdog(IN := FALSE);

			(*Kuka.PlcToKuka.bExtStart := FALSE;
			Kuka.PlcToKuka.bPgNoParity := FALSE;
			Kuka.PlcToKuka.bPgNoValid := FALSE;*)

			etKukaStart := ET_KukaStart_eWfPgNoReq;              (* Next step *)

		ELSIF Kuka.KukaToPlc.bStopMess
		THEN
			tonWatchdog(IN := FALSE);

			Kuka.PlcToKuka.bExtStart := FALSE;
			Kuka.PlcToKuka.bPgNoParity := FALSE;
			Kuka.PlcToKuka.bPgNoValid := FALSE;

			udnErrorNo := 3;                     (* Error number *)
			
			etKukaStart := ET_KukaStart_eError;              (* Next step *)

		END_IF

	ET_KukaStart_eWfPgNoReq:
		nWatchdog := nWatchdog + 1;

		IF Kuka.KukaToPlc.bPgNoReq
		     AND Kuka.KukaToPlc.bProAct
		     AND Kuka.KukaToPlc.bOnPath
		     AND NOT Kuka.KukaToPlc.bApplRun
		     AND NOT Kuka.KukaToPlc.bStopMess
		THEN
			(*Kuka.PlcToKuka.bExtStart := FALSE;
			Kuka.PlcToKuka.bPgNoParity := FALSE;
			Kuka.PlcToKuka.bPgNoValid := FALSE;*)

			nWatchdog := 0;

			etKukaStart := ET_KukaStart_ePgNoParity;              (* Next step *)

		ELSIF Kuka.KukaToPlc.bStopMess
			   OR nWatchdog > 1000
		THEN
			Kuka.PlcToKuka.bExtStart := FALSE;
			Kuka.PlcToKuka.bPgNoParity := FALSE;
			Kuka.PlcToKuka.bPgNoValid := FALSE;

			udnErrorNo := 4;                     (* Error number *)
			
			etKukaStart := ET_KukaStart_eError;              (* Next step *)

		END_IF

	ET_KukaStart_ePgNoParity:
		nWatchdog := nWatchdog + 1;

		Kuka.PlcToKuka.bPgNoParity := CHECK_PARITY(in :=  Kuka.PlcToKuka.nPgNo, p := 1);

		IF Kuka.KukaToPlc.bProAct
		     AND Kuka.KukaToPlc.bOnPath
		     AND NOT Kuka.KukaToPlc.bApplRun
		     AND NOT Kuka.KukaToPlc.bStopMess
		THEN
			nWatchdog := 0;

			etKukaStart := ET_KukaStart_ePgNoValid;              (* Next step *)

		ELSIF Kuka.KukaToPlc.bStopMess
			    OR nWatchdog > 1000
		THEN
			Kuka.PlcToKuka.bExtStart := FALSE;
			Kuka.PlcToKuka.bPgNoParity := FALSE;
			Kuka.PlcToKuka.bPgNoValid := FALSE;
			
			udnErrorNo := 5;                     (* Error number *)
			
			etKukaStart := ET_KukaStart_eError;              (* Next step *)

		END_IF

	ET_KukaStart_ePgNoValid:
		Kuka.PlcToKuka.bPgNoValid := TRUE;

		IF NOT Kuka.KukaToPlc.bPgNoReq
		     AND NOT Kuka.KukaToPlc.bInHome
		     AND NOT Kuka.KukaToPlc.arbInHome[1]
		     AND Kuka.KukaToPlc.bProAct
		     AND Kuka.KukaToPlc.bOnPath
		     AND Kuka.KukaToPlc.bApplRun
		     AND NOT Kuka.KukaToPlc.bStopMess
		THEN
			Kuka.PlcToKuka.bExtStart := FALSE;
			Kuka.PlcToKuka.bPgNoParity := FALSE;
			Kuka.PlcToKuka.bPgNoValid := FALSE;

			etKukaStart := ET_KukaStart_eWfProgFinish;              (* Next step *)

		ELSIF Kuka.KukaToPlc.bStopMess
		THEN
			Kuka.PlcToKuka.bExtStart := FALSE;
			Kuka.PlcToKuka.bPgNoParity := FALSE;
			Kuka.PlcToKuka.bPgNoValid := FALSE;

			udnErrorNo := 6;                     (* Error number *)
			
			etKukaStart := ET_KukaStart_eError;              (* Next step *)

		END_IF

	ET_KukaStart_eWfProgFinish:
		IF ((Kuka.KukaToPlc.bInHome
		      AND Kuka.PlcToKuka.nPgNo < 100)
		     OR (Kuka.PlcToKuka.nPgNo >= 100
			    AND Kuka.KukaToPlc.arbInHome[1]))
	     	    AND Kuka.KukaToPlc.bProAct
	    	    AND Kuka.KukaToPlc.bOnPath
		    AND NOT Kuka.KukaToPlc.bApplRun
	     	    AND NOT Kuka.KukaToPlc.bStopMess
		THEN
			Kuka.PlcToKuka.bExtStart := FALSE;
			Kuka.PlcToKuka.bPgNoParity := FALSE;
			Kuka.PlcToKuka.bPgNoValid := FALSE;

			etKukaStart := ET_KukaStart_eDone;              (* Next step *)

		ELSIF Kuka.KukaToPlc.bStopMess
		THEN
			Kuka.PlcToKuka.bExtStart := FALSE;
			Kuka.PlcToKuka.bPgNoParity := FALSE;
			Kuka.PlcToKuka.bPgNoValid := FALSE;

			udnErrorNo := 7;                     (* Error number *)
			
			etKukaStart := ET_KukaStart_eError;              (* Next step *)

		END_IF

	ET_KukaStart_eError:
		bBusy := FALSE;						(* Command busy *)
		bError := TRUE;						(* Command error  *)

		etKukaStart := ET_KukaStart_eNoExecute;

	ET_KukaStart_eDone:
		bDone := TRUE;						(* Command done *)
		bBusy := FALSE;						(* Command busy *)

		etKukaStart := ET_KukaStart_eNoExecute;

	ET_KukaStart_eNoExecute:
		IF NOT bStart
		THEN
			(* Reset outputs *)
			bDone := FALSE;						(* Command done *)
			bBusy := FALSE;						(* Command busy *)
			bError := FALSE;						(* Command error  *)

			nWatchdog := 0;

			Kuka.PlcToKuka.bExtStart := FALSE;
			Kuka.PlcToKuka.bPgNoParity := FALSE;
			Kuka.PlcToKuka.bPgNoValid := FALSE;

			etKukaStart := ET_KukaStart_eWaitExecute;
		END_IF
END_CASE;

END_FUNCTION_BLOCK

// ---- POUs/Tc3 Objects/ExternalHardware/KUKA/FB_KUKA_REF_1.TcPOU
FUNCTION_BLOCK FB_KUKA_REF_1
VAR_INPUT
	KukaToPlc			:ST_KUKATOPLC;
	PlcToKuka			:ST_PLCTOKUKA;
END_VAR
VAR_OUTPUT

END_VAR
VAR_IN_OUT

END_VAR
VAR

END_VAR

;

END_FUNCTION_BLOCK

// ---- POUs/Tc3 Objects/ExternalHardware/KUKA/FB_KUKA_Reset_1.TcPOU
FUNCTION_BLOCK FB_KUKA_Reset_1
(*

The function block used to reset the kuka message.

Constructor: 		Patryk Panylo
Company:		E. Riexinger GmbH
Date:			18.11.2016
Version:			1.00

Date:			Revision:		Who:				Comment

*)
VAR_INPUT
	(* Input variables / Eingang Variablen *)
	bReset						:BOOL;		(* Execut the function block *)
	bExtReset					:BOOL;
END_VAR
VAR_OUTPUT
	(* Output variables / Ausgang Variablen *)
	bDone						:BOOL;			(* Status = TRUE indicates that the axis is ready for operation. *)
	bError						:BOOL;			(* Error *)
	udnErrorNo					:UDINT;			(* Error number *)
	sErrorMsg					:STRING; 		(* Error message *)
END_VAR
VAR_IN_OUT
	(* Input Output variables / Ausgang Variablen *)
	Kuka						:ST_KUKA_REF;
END_VAR
VAR
	(* Enummerations *)

	(* Variables *)

	(* References *)

	(* Interfaces *)

	(* Instances *)
	rtExecute						:R_TRIG;
	rtExtReset					:R_TRIG;
	rtDrivesOk					:R_TRIG;
	tonConfMess					:TON;
END_VAR


rtExecute(CLK := bReset);
rtExtReset(CLK := bExtReset
			       AND Kuka.KukaToPlc.bStopMess);
rtDrivesOk(CLK := Kuka.KukaToPlc.bPeriRdy
	   		        AND Kuka.PlcToKuka.bDrivesOff
			        AND Kuka.KukaToPlc.bStopMess);

tonConfMess(
	IN := Kuka.PlcToKuka.bConfMess,
	PT := t#100ms
);

IF rtExecute.Q
     OR rtExtReset.Q
     OR rtDrivesOk.Q
THEN
	Kuka.PlcToKuka.bConfMess := TRUE;

ELSIF tonConfMess.Q
	   OR NOT Kuka.KukaToPlc.bStopMess
THEN
	Kuka.PlcToKuka.bConfMess := FALSE;
END_IF;
(*
IF NOT Kuka.KukaToPlc.bStopMess       (* Error *)
THEN
	Kuka.PlcToKuka.bConfMess := FALSE;
END_IF;
*)

bDone := bReset
		AND NOT Kuka.KukaToPlc.bStopMess;        (* Error *)

END_FUNCTION_BLOCK

// ---- POUs/Tc3 Objects/ExternalHardware/KUKA/FB_KUKA_StartProg_1.TcPOU
FUNCTION_BLOCK FB_KUKA_StartProg_1
(*

The function block used to start kuka

Constructor: 		Patryk Panylo
Company:		E. Riexinger GmbH
Date:			18.11.2016
Version:			1.00

Date:			Revision:		Who:				Comment

*)
VAR_INPUT
	(* Input variables / Eingang Variablen *)
	bEnable						:BOOL;			(* Signal FB enable *)
	bStart						:BOOL;			(* Execute start *)
	nProgNo						:INT;			(* Program number *)
	tMaxRefTime					:TIME := t#60s;	(* Maximal referenc time *)
END_VAR
VAR_OUTPUT
	(* Output variables / Ausgang Variablen *)
	bRunning					:BOOL;						(* Program running *)
	bDone						:BOOL;						(* Program done *)
	bBusy						:BOOL;						(* Program busy *)
	bError						:BOOL;						(* Error *)
	udnErrorNo					:UDINT;
END_VAR
VAR_IN_OUT
	(* Input Output variables / Ausgang Variablen *)
	Kuka						:ST_KUKA_REF;
END_VAR
VAR
	(* Enummerations *)
	etKukaStart					:ET_KukaStart;

	(* Variables *)
	bFirstTime					:BOOL;

	nWatchdog					:INT;

	(* References *)

	(* Interfaces *)

	(* Instances *)
	rtStart						:R_TRIG;
	tonWatchdog					:TON;

END_VAR


IF NOT bEnable
THEN
	bDone := FALSE;					(* Program done *)
	bBusy := FALSE;                                  	(* Program not busy *)
	bError := FALSE;                                 	(* Program not error *)
	udnErrorNo := 0;                                 		(* Error number *)

	Kuka.PlcToKuka.bExtStart := FALSE;
	Kuka.PlcToKuka.bPgNoParity := FALSE;
	Kuka.PlcToKuka.bPgNoValid := FALSE;

	RETURN;
END_IF;

IF NOT bFirstTime
THEN
	tonWatchdog(IN := FALSE);

	Kuka.PlcToKuka.bExtStart := FALSE;
	Kuka.PlcToKuka.bPgNoParity := FALSE;
	Kuka.PlcToKuka.bPgNoValid := FALSE;

	etKukaStart := ET_KukaStart_eWaitExecute;              (* Next step *)

	bFirstTime := TRUE;
END_IF

bRunning := Kuka.KukaToPlc.bApplRun
		      AND Kuka.KukaToPlc.bProAct;

IF NOT Kuka.PlcToKuka.bDrivesOff
     OR NOT Kuka.PlcToKuka.bMoveEnable
     OR NOT Kuka.KukaToPlc.bUserSafe
     OR NOT Kuka.KukaToPlc.bAlarmStop
     OR NOT Kuka.KukaToPlc.bPeriRdy
     OR Kuka.PlcToKuka.bDrivesOn
     OR Kuka.KukaToPlc.bStopMess
THEN
	Kuka.PlcToKuka.bExtStart := FALSE;
	Kuka.PlcToKuka.bPgNoParity := FALSE;
	Kuka.PlcToKuka.bPgNoValid := FALSE;

	etKukaStart := ET_KukaStart_eWaitExecute;              (* Next step *)

	RETURN;
END_IF

(* Wait for triger *)
rtStart(
	CLK := bStart
);

IF rtStart.Q
    AND NOT Kuka.KukaToPlc.bProAct
THEN
	etKukaStart := ET_KukaStart_eWaitExecute;              (* Next step *)

END_IF

(* Send command *)
CASE etKukaStart OF

	ET_KukaStart_eWaitExecute:
		bBusy := FALSE;                                     	(* Program not busy *)
		bError := FALSE;                         		(* Program not error *)
		udnErrorNo := 0;                         		(* Error number *)

		IF rtStart.Q
		THEN
			nWatchdog := 0;
			bDone:= FALSE;                               		(* Program done *)
			bBusy := TRUE;                                  	(* Program busy *)

			tonWatchdog(IN := FALSE);

			Kuka.PlcToKuka.bExtStart := FALSE;
			Kuka.PlcToKuka.bPgNoParity := FALSE;
			Kuka.PlcToKuka.bPgNoValid := FALSE;
			Kuka.PlcToKuka.nPgNo := nProgNo;

			etKukaStart := ET_KukaStart_eExtStart;              (* Next step *)

		END_IF

	ET_KukaStart_eExtStart:
		nWatchdog := nWatchdog + 1;

		Kuka.PlcToKuka.bExtStart := TRUE;
		Kuka.PlcToKuka.bPgNoParity := FALSE;
		Kuka.PlcToKuka.bPgNoValid := FALSE;

		IF Kuka.KukaToPlc.bProAct
		     AND Kuka.KukaToPlc.bOnPath
		     AND NOT Kuka.KukaToPlc.bStopMess
		THEN
			nWatchdog := 0;

			Kuka.PlcToKuka.bExtStart := FALSE;
			Kuka.PlcToKuka.bPgNoParity := FALSE;
			Kuka.PlcToKuka.bPgNoValid := FALSE;

			etKukaStart := ET_KukaStart_eWfInHome;              (* Next step *)

		ELSIF Kuka.KukaToPlc.bStopMess
			    OR nWatchdog > 1000
		THEN
			Kuka.PlcToKuka.bExtStart := FALSE;
			Kuka.PlcToKuka.bPgNoParity := FALSE;
			Kuka.PlcToKuka.bPgNoValid := FALSE;
			
			udnErrorNo := 1;                     (* Error number *)
			
			etKukaStart := ET_KukaStart_eError;              (* Next step *)

		END_IF

	ET_KukaStart_eWfInHome:
		tonWatchdog(
			IN := Kuka.PlcToKuka.nOverride > 0,
			PT:= tMaxRefTime
		);

		IF tonWatchdog.Q
		THEN
			tonWatchdog(IN := FALSE);

			Kuka.PlcToKuka.bExtStart := FALSE;
			Kuka.PlcToKuka.bPgNoParity := FALSE;
			Kuka.PlcToKuka.bPgNoValid := FALSE;

			udnErrorNo := 2;

			etKukaStart := ET_KukaStart_eError;             (* Next step *)

		ELSIF Kuka.KukaToPlc.bInHome
		     	    AND Kuka.KukaToPlc.bProAct
		    	    AND Kuka.KukaToPlc.bOnPath
		     	    AND NOT Kuka.KukaToPlc.bStopMess
		THEN
			tonWatchdog(IN := FALSE);

			Kuka.PlcToKuka.bExtStart := FALSE;
			Kuka.PlcToKuka.bPgNoParity := FALSE;
			Kuka.PlcToKuka.bPgNoValid := FALSE;

			etKukaStart := ET_KukaStart_eWfPgNoReq;              (* Next step *)

		ELSIF Kuka.KukaToPlc.bStopMess
		THEN
			tonWatchdog(IN := FALSE);

			Kuka.PlcToKuka.bExtStart := FALSE;
			Kuka.PlcToKuka.bPgNoParity := FALSE;
			Kuka.PlcToKuka.bPgNoValid := FALSE;

			udnErrorNo := 3;                     (* Error number *)
			
			etKukaStart := ET_KukaStart_eError;              (* Next step *)

		END_IF

	ET_KukaStart_eWfPgNoReq:
		nWatchdog := nWatchdog + 1;

		IF Kuka.KukaToPlc.bPgNoReq
		     AND Kuka.KukaToPlc.bProAct
		     AND Kuka.KukaToPlc.bOnPath
		     AND NOT Kuka.KukaToPlc.bStopMess
		THEN
			Kuka.PlcToKuka.bExtStart := FALSE;
			Kuka.PlcToKuka.bPgNoParity := FALSE;
			Kuka.PlcToKuka.bPgNoValid := FALSE;

			nWatchdog := 0;

			etKukaStart := ET_KukaStart_ePgNoParity;              (* Next step *)

		ELSIF Kuka.KukaToPlc.bStopMess
			   OR nWatchdog > 1000
		THEN
			Kuka.PlcToKuka.bExtStart := FALSE;
			Kuka.PlcToKuka.bPgNoParity := FALSE;
			Kuka.PlcToKuka.bPgNoValid := FALSE;

			udnErrorNo := 4;                     (* Error number *)
			
			etKukaStart := ET_KukaStart_eError;              (* Next step *)

		END_IF

	ET_KukaStart_ePgNoParity:
		nWatchdog := nWatchdog + 1;

		Kuka.PlcToKuka.bPgNoParity := CHECK_PARITY(in :=  Kuka.PlcToKuka.nPgNo, p := 1);

		IF Kuka.KukaToPlc.bProAct
		     AND Kuka.KukaToPlc.bOnPath
		     AND NOT Kuka.KukaToPlc.bStopMess
		THEN
			nWatchdog := 0;

			etKukaStart := ET_KukaStart_ePgNoValid;              (* Next step *)

		ELSIF Kuka.KukaToPlc.bStopMess
			    OR nWatchdog > 1000
		THEN
			Kuka.PlcToKuka.bExtStart := FALSE;
			Kuka.PlcToKuka.bPgNoParity := FALSE;
			Kuka.PlcToKuka.bPgNoValid := FALSE;
			
			udnErrorNo := 5;                     (* Error number *)
			
			etKukaStart := ET_KukaStart_eError;              (* Next step *)

		END_IF

	ET_KukaStart_ePgNoValid:
		Kuka.PlcToKuka.bPgNoValid := TRUE;

		IF NOT Kuka.KukaToPlc.bPgNoReq
		     AND NOT Kuka.KukaToPlc.bInHome
		     AND Kuka.KukaToPlc.bProAct
		     AND Kuka.KukaToPlc.bOnPath
		     AND NOT Kuka.KukaToPlc.bStopMess
		THEN
			Kuka.PlcToKuka.bExtStart := FALSE;
			Kuka.PlcToKuka.bPgNoParity := FALSE;
			Kuka.PlcToKuka.bPgNoValid := FALSE;

			etKukaStart := ET_KukaStart_eWfProgFinish;              (* Next step *)

		ELSIF Kuka.KukaToPlc.bStopMess
		THEN
			Kuka.PlcToKuka.bExtStart := FALSE;
			Kuka.PlcToKuka.bPgNoParity := FALSE;
			Kuka.PlcToKuka.bPgNoValid := FALSE;

			udnErrorNo := 6;                     (* Error number *)
			
			etKukaStart := ET_KukaStart_eError;              (* Next step *)

		END_IF

	ET_KukaStart_eWfProgFinish:
		IF Kuka.KukaToPlc.bInHome
	     	    AND Kuka.KukaToPlc.bProAct
	    	    AND Kuka.KukaToPlc.bOnPath
	     	    AND NOT Kuka.KukaToPlc.bStopMess
		THEN
			Kuka.PlcToKuka.bExtStart := FALSE;
			Kuka.PlcToKuka.bPgNoParity := FALSE;
			Kuka.PlcToKuka.bPgNoValid := FALSE;

			etKukaStart := ET_KukaStart_eDone;              (* Next step *)

		ELSIF Kuka.KukaToPlc.bStopMess
		THEN
			Kuka.PlcToKuka.bExtStart := FALSE;
			Kuka.PlcToKuka.bPgNoParity := FALSE;
			Kuka.PlcToKuka.bPgNoValid := FALSE;

			udnErrorNo := 7;                     (* Error number *)
			
			etKukaStart := ET_KukaStart_eError;              (* Next step *)

		END_IF

	ET_KukaStart_eError:
		bBusy := FALSE;						(* Command busy *)
		bError := TRUE;						(* Command error  *)

		etKukaStart := ET_KukaStart_eNoExecute;

	ET_KukaStart_eDone:
		bDone := TRUE;						(* Command done *)
		bBusy := FALSE;						(* Command busy *)

		etKukaStart := ET_KukaStart_eNoExecute;

	ET_KukaStart_eNoExecute:
		IF NOT bStart
		THEN
			(* Reset outputs *)
			bDone := FALSE;						(* Command done *)
			bBusy := FALSE;						(* Command busy *)
			bError := FALSE;						(* Command error  *)

			nWatchdog := 0;

			Kuka.PlcToKuka.bExtStart := FALSE;
			Kuka.PlcToKuka.bPgNoParity := FALSE;
			Kuka.PlcToKuka.bPgNoValid := FALSE;

			etKukaStart := ET_KukaStart_eWaitExecute;
		END_IF
END_CASE;

END_FUNCTION_BLOCK

// ---- POUs/Tc3 Objects/ExternalHardware/KUKA/FB_MoveToKukaRef_1.TcPOU
FUNCTION_BLOCK FB_MoveToKukaRef_1
VAR_INPUT
	stRobotToPlc					:ST_ROBOTTOPLC;
END_VAR
VAR_OUTPUT
	stPlcToRobot					:ST_PLCTOROBOT;
END_VAR
VAR_IN_OUT
	Kuka						:ST_KUKA_REF;				(* The KUKA_REF data type  is an interface between the PLC and the KUKA and contains axis information *)
END_VAR
VAR
	rtForceToBase				:R_TRIG;
	rtForceToWork				:R_TRIG;
	rtCutoffToBase				:R_TRIG;
	rtCutoffToWork				:R_TRIG;

	rtMEStartHeat					:R_TRIG;
	rtMEStopHeat				:R_TRIG;
	rtMEStartExtruding				:R_TRIG;
	rtMEStopExtruding				:R_TRIG;
	rtMEStartFlush				:R_TRIG;
	rtMEStopFlush				:R_TRIG;
END_VAR


(* Set general parameter *)


(* Copy the actual values from the robot to the kuka reference *)
Kuka.KukaToPlc.bPgNoReq := stRobotToPlc.arbyInput[2].0;						(* $OUT[33] - A change of signal requests the higher-level controller to send a program number / PGNO Req-Signalwechsel fordert Leitrechner Programmnr. zu senden *)

Kuka.KukaToPlc.bApplRun := stRobotToPlc.arbyInput[2].1;						(* $OUT[34] - Program is currently being executed / TRUE wenn Programm abgearbeitet wird *)
Kuka.KukaToPlc.bErrToPlc := stRobotToPlc.arbyInput[2].2;						(* $OUT[35] - Error output to PLC / Steuerungs- oder Technologiefehler aufgetreten *)
Kuka.KukaToPlc.bInWorkArea := stRobotToPlc.arbyInput[2].3;					(* $OUT[36] - Robot in work area / Roboter in Bearbeitunsbereich*)

Kuka.KukaToPlc.bIOActConf := stRobotToPlc.arbyInput[0].0;						(* $OUT[140] - This output is TRUE if Automatic External mode is selected and the input $I_O_ACT is TRUE. / *)
Kuka.KukaToPlc.bT1:= stRobotToPlc.arbyInput[0].1;							(* $OUT[993] - Operating mode T1 / Betriebsart T1 *)
Kuka.KukaToPlc.bT2 := stRobotToPlc.arbyInput[0].2;							(* $OUT[994] - Operating mode T2/ Betriebsart T2 *)
Kuka.KukaToPlc.bAut := stRobotToPlc.arbyInput[0].3;							(* $OUT[995] - Operating mode Aut / Betriebsart Aut *)
Kuka.KukaToPlc.bExt := stRobotToPlc.arbyInput[0].4;							(* $OUT[996] - Operating mode Ext / Betriebsart Ext *)
Kuka.KukaToPlc.bOnPath := stRobotToPlc.arbyInput[0].5;						(* $OUT[997] - Set as long as the robot stays on its programmed path / TRUE solange sich Rob. auf programmierten Bahn befindet *)
Kuka.KukaToPlc.bInHome := stRobotToPlc.arbyInput[0].6;						(* $OUT[1000] - Whether or not the robot is in its HOME position  / In Home Position *)
Kuka.KukaToPlc.bStopMess := stRobotToPlc.arbyInput[0].7; 						(* $OUT[1010] - Any message occurring which requires the robot to be stopped / Störung Roboter *)
Kuka.KukaToPlc.bUserSafe := stRobotToPlc.arbyInput[1].0;						(* $OUT[1011] - If the safety fence monitoring switch is opened (AUT mode) or an enabling switch is released (T1 or T2 mode). / Abfrage Schutzgitter(Auto)/Zustimmungsschalter(Test) *)
Kuka.KukaToPlc.bPeriRdy := stRobotToPlc.arbyInput[1].1;						(* $OUT[1012] - Robot drives are switched on / TRUE wenn Roboterantriebe eingeschaltet *)
Kuka.KukaToPlc.bAlarmStop := stRobotToPlc.arbyInput[1].2;						(* $OUT[1013] - Emergency stop / Not Aus *)
Kuka.KukaToPlc.bProAct := stRobotToPlc.arbyInput[1].3;							(* $OUT[1021] - Whenever a process is active / Programmbearbeitung aktiv *)

Kuka.KukaToPlc.arbInHome[1]:= stRobotToPlc.arbyInput[3].1;					(* $OUT[1003] - Whether or not the robot is in its HOME position  / In Home Position *)
Kuka.KukaToPlc.arbInHome[2] := stRobotToPlc.arbyInput[3].2;					(* $OUT[1004] - Whether or not the robot is in its HOME position  / In Home Position *)
Kuka.KukaToPlc.arbInHome[3] := stRobotToPlc.arbyInput[3].3;					(* $OUT[1005] - Whether or not the robot is in its HOME position  / In Home Position *)
Kuka.KukaToPlc.arbInHome[4] := stRobotToPlc.arbyInput[3].4;					(* $OUT[1006] - Whether or not the robot is in its HOME position  / In Home Position *)
Kuka.KukaToPlc.arbInHome[5] := stRobotToPlc.arbyInput[3].5;					(* $OUT[1007] - Whether or not the robot is in its HOME position  / In Home Position *)

rtForceToBase(CLK := stRobotToPlc.arbyInput[12].0); Kuka.KukaToPlc.bForceToBase := rtForceToBase.Q;					(* $OUT[10] - Move force to base position *)
rtForceToWork(CLK := stRobotToPlc.arbyInput[12].1); Kuka.KukaToPlc.bForceToWork := rtForceToWork.Q;					(* $OUT[11] - Move force to work position *)
rtCutoffToBase(CLK := stRobotToPlc.arbyInput[12].2); Kuka.KukaToPlc.bCutoffToBase := rtCutoffToBase.Q;					(* $OUT[12] - Move cutoff to base position *)
rtCutoffToWork(CLK := stRobotToPlc.arbyInput[12].3); Kuka.KukaToPlc.bCutoffToWork := rtCutoffToWork.Q;					(* $OUT[13] - Move cutoffe to work position *)

rtMEStartHeat(CLK := stRobotToPlc.arbyInput[13].0); Kuka.KukaToPlc.bMEStartHeat := rtMEStartHeat.Q;						(* $OUT[18] - Start heat *)
rtMEStopHeat(CLK := stRobotToPlc.arbyInput[13].1); Kuka.KukaToPlc.bMEStopHeat := rtMEStopHeat.Q;						(* $OUT[19] - Stop heat *)
rtMEStartExtruding(CLK := stRobotToPlc.arbyInput[13].2); Kuka.KukaToPlc.bMEStartExtruding := rtMEStartExtruding.Q;			(* $OUT[20] - Start extruding *)
rtMEStopExtruding(CLK := stRobotToPlc.arbyInput[13].3); Kuka.KukaToPlc.bMEStopExtruding := rtMEStopExtruding.Q;			(* $OUT[21] - Stop extruding *)
rtMEStartFlush(CLK := stRobotToPlc.arbyInput[13].4); Kuka.KukaToPlc.bMEStartFlush := rtMEStartFlush.Q;					(* $OUT[22] - Start flush *)
rtMEStopFlush(CLK := stRobotToPlc.arbyInput[13].5); Kuka.KukaToPlc.bMEStopFlush := rtMEStopFlush.Q;					(* $OUT[23] - Stop flush *)
Kuka.KukaToPlc.nMEExtrudingSpeed := BYTE_TO_INT(stRobotToPlc.arbyInput[10]);	(* $OUT[100] - Extruding speed [%] *)

(* Copy the setpoint values from the kuka reference to the robot *)
stPlcToRobot.arbyOutput[4] := INT_TO_BYTE(Kuka.PlcToKuka.nPgNo);		(* $IN[33] - Program number / Programmnummer *)
																	(* $IN[33]  + 8 = $IN[41], PGNO_LENGTH = 8 (max. 16) *)
stPlcToRobot.arbyOutput[2].0 := Kuka.PlcToKuka.bPgNoParity;				(* $IN[41] - Input to which the parity bit is transferred from the higher-level controller / Übertragen des Paritätsbit vom Leitrechner *)
stPlcToRobot.arbyOutput[2].1 := Kuka.PlcToKuka.bPgNoValid;				(* $IN[42] - Input to which the command to read the program number is transferred from the higher-level controller / Einlesen der Programmnumer vom Leitrechener *)

stPlcToRobot.arbyOutput[0].0 := Kuka.PlcToKuka.bDrivesOn;					(* $IN[140] - Switch on the robot drives / Einschalten der Roboterantriebe *)
stPlcToRobot.arbyOutput[0].1 := Kuka.PlcToKuka.bDrivesOff;					(* $IN[141] - Switch off the robot drives / Abschalten der Roboterantriebe *)
stPlcToRobot.arbyOutput[0].2 := Kuka.PlcToKuka.bMoveEnable;				(* $IN[143] - Check the robot drives. TRUE Jogging and program execution are possible / Kontrolle der Roboterantriebe *)
stPlcToRobot.arbyOutput[0].3 := Kuka.PlcToKuka.bIOAct;					(* $IN[1025] - If this input is TRUE, the Automatic External interface is active. Default setting:$IN[1025]. *)
stPlcToRobot.arbyOutput[0].4 := Kuka.PlcToKuka.bConfMess;				(* $IN[142] - Acknowledge error / Quittieren von Fehlermeldungen durch den Leitrechner *)
stPlcToRobot.arbyOutput[0].5 := Kuka.PlcToKuka.bExtStart;					(* $IN[145] - If the I/O interface is active, this input can be set to start or continue a program / Extern Start *)

stPlcToRobot.arbyOutput[0].6 := Kuka.PlcToKuka.bCheckMovena;			(* TRUE MOVE_ENABLE monitoring is activated / Überwachung für MOVE_ENABLE *)

stPlcToRobot.arbyOutput[1].0 := Kuka.PlcToKuka.bPgReset;					(* $IN[148] - Cancel a program / Programm abbrechen *)

stPlcToRobot.arbyOutput[10] := INT_TO_BYTE(Kuka.PlcToKuka.nOverride);	(* $IN[100] - Override *)

stPlcToRobot.arbyOutput[6] := INT_TO_BYTE(Kuka.PlcToKuka.nCutOffDist);						(* $IN[50] - Distance of cutoff *)
stPlcToRobot.arbyOutput[7] := INT_TO_BYTE(SHR(Kuka.PlcToKuka.nCutOffDist,8));

stPlcToRobot.arbyOutput[8] := INT_TO_BYTE(Kuka.PlcToKuka.nExtruderOffDist);					(* $IN[66] - Distance aftre extruder is off *)
stPlcToRobot.arbyOutput[9] := INT_TO_BYTE(SHR(Kuka.PlcToKuka.nExtruderOffDist,8));

stPlcToRobot.arbyOutput[14] := UINT_TO_BYTE(Kuka.PlcToKuka.unExtruderStartTime);				(* $IN[82] - Extruder start time *)
stPlcToRobot.arbyOutput[15] := UINT_TO_BYTE(SHR(Kuka.PlcToKuka.unExtruderStartTime,8));

stPlcToRobot.arbyOutput[12].0 := Kuka.PlcToKuka.bForceInBase;			(* $IN[10] - Force in base position *)
stPlcToRobot.arbyOutput[12].1 := Kuka.PlcToKuka.bForceInWork;			(* $IN[11] - Force in work position *)
stPlcToRobot.arbyOutput[12].2 := Kuka.PlcToKuka.bCutoffInBase;			(* $IN[12] - Cutoff in base position *)
stPlcToRobot.arbyOutput[12].3 := Kuka.PlcToKuka.bCutoffInWork;			(* $IN[13] - Cutoff in work position *)

stPlcToRobot.arbyOutput[13].0 := Kuka.PlcToKuka.bMEHeat;				(* $IN[18] - Heat status ON = TRUE, OFF = FALSE *)
stPlcToRobot.arbyOutput[13].1 := Kuka.PlcToKuka.bMEHeating;			(* $IN[19] - Heating status ON = TRUE, OFF = FALSE *)
stPlcToRobot.arbyOutput[13].2 := Kuka.PlcToKuka.bMEHeated;			(* $IN[20] - Heated status ON = TRUE, OFF = FALSE *)
stPlcToRobot.arbyOutput[13].3 := Kuka.PlcToKuka.bMEExtruding;			(* $IN[21] - Extruder status ON = TRUE, OFF = FALSE *)

END_FUNCTION_BLOCK

// ---- POUs/Tc3 Objects/ExternalHardware/Munsch/FB_MunschExtruderAir_1.TcPOU
FUNCTION_BLOCK FB_MunschExtruderAir_1
(*

The function block used to control air pressure.

Constructor: 		Patryk Panylo
Company:		E. Riexinger GmbH
Date:			04.11.2016
Version:			1.00

Date:			Revision:		Who:				Comment
dd.mm.yyyy		x.xx			Initials			comment

*)
VAR_INPUT
	(* Input variables / Eingang Variablen *)
	bEnable					:BOOL;						(* Enable FB signal *)
	bIn						:BOOL;						(* Input signal *)
	bExtruderAirOn			:BOOL;						(* Extruder air on *)
	tAirOk					:TIME := t#5s;					(* Timer to delay output air ok *)
	tAirOff					:TIME := t#5s;					(* Timer to delay output air off *)
	tTimeOut					:TIME := t#5s;					(* Timeout *)
END_VAR
VAR_OUTPUT
	(* Output variables / Ausgang Variablen *)
	bAirOk					:BOOL;						(* Air pressure ok *)
	bAirOn					:BOOL;						(* Air pressure on *)
	bError					:BOOL;						(* Error by no air pressure *)
	udnErrorNo				:UDINT;
	udnMessageNo			:UDINT;
END_VAR
VAR
	(* Enummerations *)

	(* Variables *)

	(* References *)

	(* Interfaces *)

	(* Instances *)
	tonDelayAirOk				:TON;						(* Timer to delay *)
	tofDelayAirOff					:TOF;						(* Timer to delay *)
	fbExtrudingAir					:FB_AirPressure;
END_VAR


IF NOT bEnable
THEN
	fbExtrudingAir(
		bEnable := FALSE
	);

	bAirOk := FALSE;
	RETURN;
END_IF

fbExtrudingAir(
	bEnable := bEnable,
	bIn := bIn,
	bNoEStop := bExtruderAirOn,
	tTimeOut := tTimeOut,
	bError => bError,
	udnErrorNo => udnErrorNo,
	udnMessageNo => udnMessageNo
);

tonDelayAirOk(
	IN := fbExtrudingAir.bOut,
	PT := tAirOk
);

bAirOk := tonDelayAirOk.Q;

tofDelayAirOff(
	IN := fbExtrudingAir.bAirOn,
	PT := tAirOff
);

bAirOn := tofDelayAirOff.Q;

END_FUNCTION_BLOCK

// ---- POUs/Tc3 Objects/ExternalHardware/Munsch/FB_MunschExtruder_1.TcPOU
FUNCTION_BLOCK FB_MunschExtruder_1
(*

This function block is used to send and recive data's via KL600x to/from Munsch extruder.

KL600x configuration is 	1200 8-N-1

Constructor: 		Patryk Panylo
Company:		E. Riexinger GmbH
Date:			14.09.2016
Version:			1.00

Date:			Revision:		Who:				Comment
dd.mm.yyyy		x.xx			Initials			comment

*)
VAR_INPUT
	(* Input variables / Eingang Variablen *)
	bEnable						:BOOL;					(* Enable FB *)
	sDeviceNetId					:STRING;				(* Fieldbus master NetId *)
	unSlaveAddr 					:UINT;					(* Fixed address of the slave *)
	sDateTime					:STRING;				(* Current date and time *)
	bReset						:BOOL;					(* Reset *)
	bSendExe					:BOOL;					(* Send execute *)
	tSendPeriod					:TIME := t#0s;				(* Send data every period. If tSendPeriod is 0 then th function is not active *)
	stMunschCmd				:ST_MUNSCH_CMD_Data;
	tTimeOut 					:TIME := t#2s;				(* Timout  *)
END_VAR
VAR_OUTPUT
	(* Output variables / Ausgang Variablen *)
	stMunschRes					:ST_MUNSCH_RES_Data;
	bInterfaceReady				:BOOL;				(* Interface ready to use *)
	bInterfaceError				:BOOL;				(* Interface error *)
	bStringReceived				:BOOL;				(* String received *)
END_VAR
VAR_IN_OUT
	(* Input Output variables / Ausgang Variablen *)
	stRXbuffer 					:ComBuffer;
	stTXbuffer					:ComBuffer;
END_VAR
VAR
	(* Enummerations *)

	(* Variables *)
	sSendString					:STRING;
	sReceivedString				:STRING;

	bFirstTime					:BOOL;					(* First PLC cycle *)

	(* References *)

	(* Interfaces *)

	(* Instances *)
	fbKL600x						:FB_KL600xData;

END_VAR
VAR CONSTANT
	bEnableRTSCTS				:BOOL := FALSE;
	udnBaudrate					:UDINT := 1200;
	unDataBits					:UINT := 8;
	sParity						:STRING := 'N';
	unStopBits					:UINT := 1;
	sStringPrefix					:STRING := '$FC';
	sStringSuffix					:STRING := '';
	byEnRTSCTSSubIndex		:BYTE := 16#01;					(* Subindex of object *)
	wEnRTSCTSIndex			:WORD := 16#8000;                 			 (* Index of object *)
	byBaudrateSubIndex			:BYTE := 16#11;					(* Subindex of object *)
	wBaudrateIndex				:WORD := 16#8000;				(* Index of object *)
	byDataFrameSubIndex			:BYTE := 16#15;					(* Subindex of object *)
	wDataFrameIndex				:WORD := 16#8000;                                     (* Index of object *)
END_VAR


IF NOT bEnable							(* Enable FB *)
THEN
	fbKL600x(
		bEnable := FALSE,
		tTimeOut:= tTimeOut,
		sReceivedString := sReceivedString,
		stRXbuffer := stRXbuffer,
		stTXbuffer := stTXbuffer
	);

	bFirstTime := FALSE;					(* First PLC cycle *)
	RETURN;
END_IF

IF NOT bFirstTime
THEN


	bFirstTime := TRUE;
END_IF

IF bReset
     AND bInterfaceError
THEN
	bInterfaceError := FALSE;
END_IF

sSendString := F_MunschCMD(
	stMunschCmd := stMunschCmd
);

fbKL600x(
	bEnable := TRUE,
	sDeviceNetId:= sDeviceNetId,
	unSlaveAddr:= unSlaveAddr,
	sDateTime:= sDateTime,
	bEnableRTSCTS := bEnableRTSCTS,
	udnBaudrate:= udnBaudrate,
	unDataBits:= unDataBits,
	sParity:= sParity,
	unStopBits:= unStopBits,
	sStringPrefix := sStringPrefix,
	sStringSuffix := sStringSuffix,
	bReset := bReset,
	bSendExe:= bSendExe,
	tSendPeriod:= tSendPeriod,
	sSendString:= sSendString,
	byEnRTSCTSSubIndex := byEnRTSCTSSubIndex,
	wEnRTSCTSIndex := wEnRTSCTSIndex,
	byBaudrateSubIndex := byBaudrateSubIndex,
	wBaudrateIndex := wBaudrateIndex,
	byDataFrameSubIndex	 := byDataFrameSubIndex,
	wDataFrameIndex := wDataFrameIndex,
	tTimeOut:= tTimeOut,
	sReceivedString := sReceivedString,
	stRXbuffer := stRXbuffer,
	stTXbuffer := stTXbuffer,
	bKL600xReady => bInterfaceReady,
	bStringReceived => bStringReceived
 );

stMunschRes := F_MunschRES(
	sResponse := sReceivedString
);

IF fbKL600x.arbError[0]
     OR fbKL600x.arbError[1]
     OR fbKL600x.arbError[2]
     OR (bStringReceived AND stMunschRes.etResponse = ET_MUNSCH_RES_CMDERROR)
THEN
	bInterfaceError := TRUE;
END_IF

END_FUNCTION_BLOCK

// ---- POUs/Tc3 Objects/ExternalHardware/Munsch/FB_MunschExtruder_AirTemp_1.TcPOU
FUNCTION_BLOCK FB_MunschExtruder_AirTemp_1
(*

The function block used to control set material temperature on munschs extruder

Constructor: 		Patryk Panylo
Company:		E. Riexinger GmbH
Date:			18.10.2015
Version:			1.00

Date:			Revision:		Who:				Comment
dd.mm.yyyy		x.xx			Initials			comment

*)
VAR_INPUT
	(* Input variables / Eingang Variablen *)
	bEnable						:BOOL;						(* Enable FB signal *)
	bExecute					:BOOL;						(* Execut the function block *)
	nAirTemp					:INT;						(* Air temperatur *)
	nMinAirTemp					:INT;						(* Minimal air temperatur *)
	nMaxAirTemp				:INT;						(* Maximal air temperatur *)
	nAirTempTolerance			:INT := 5;						(* Air temperatur tolerance*)
END_VAR
VAR_OUTPUT
	(* Output variables / Ausgang Variablen *)
	bAirTempAlarm				:BOOL;						(* Exceeded air temperature tolerance  *)
	bDone						:BOOL;						(* Program done *)
	bBusy						:BOOL;						(* Program busy *)
	bError						:BOOL;						(* Error *)
	udnErrorNo					:UDINT;
END_VAR
VAR_IN_OUT
	(* Input Output variables / Ausgang Variablen *)
	Munsch						:ST_MUNSCH_REF;
END_VAR
VAR
	(* Enummerations *)
	etMunschExtruder				:ET_MunschExtruder;

	(* Variables *)
	nWatchdog					:INT;

	(* References *)

	(* Interfaces *)

	(* Instances *)
	rtExecute						:R_TRIG;

END_VAR

IF NOT bEnable
THEN
	bDone := FALSE;					(* Program done *)
	bBusy := FALSE;                                  	(* Program not busy *)
	bError := FALSE;                                 	(* Program not error *)
	udnErrorNo := 0;                                 		(* Error number *)

	RETURN;
END_IF;

(* Wait for triger *)
rtExecute(CLK := bExecute);

(* Send command *)
CASE etMunschExtruder OF

	ET_MunschExtruder_eWaitExecute:
		IF rtExecute.Q
		THEN
			nWatchdog := 0;

			Munsch.bSetAirTemp := TRUE;
			Munsch.bSetMaterialTemp := FALSE;
			Munsch.bStartHeat := FALSE;
			Munsch.bStopHeat  := FALSE;
			Munsch.bStartExtruding := FALSE;
			Munsch.bStopExtruding  := FALSE;
			Munsch.bReadStatus := FALSE;

			etMunschExtruder := ET_MunschExtruder_eChkInterface;              (* Next step *)
		END_IF

	ET_MunschExtruder_eChkInterface:
		nWatchdog := nWatchdog + 1;

		IF NOT Munsch.bLockedInterface
		THEN
			bBusy := FALSE;                                     	(* Program not busy *)
			bError := FALSE;                         		(* Program not error *)
			udnErrorNo := 0;                         		(* Error number *)

			IF Munsch.bSetAirTemp
			THEN
				nWatchdog := 0;
				bDone:= FALSE;                               		(* Program done *)
				bBusy := TRUE;                                  	(* Program busy *)
	
				Munsch.bLockedInterface := TRUE;
				Munsch.bSendExe := FALSE;
	
				IF nAirTemp >= nMinAirTemp
				     AND nAirTemp <= nMaxAirTemp
				THEN
					etMunschExtruder := ET_MunschExtruder_eSetCMD;              (* Next step *)
				ELSE
					udnErrorNo := 1;
	
					etMunschExtruder := ET_MunschExtruder_eError;              (* Next step *)
				END_IF

			ELSE
				etMunschExtruder := ET_MunschExtruder_eError;             (* Next step *)
			END_IF

			Munsch.bSetAirTemp := FALSE;

		ELSIF nWatchdog > 1000
		THEN
			Munsch.bSetAirTemp := FALSE;

			etMunschExtruder := ET_MunschExtruder_eError;             (* Next step *)
		END_IF

	ET_MunschExtruder_eSetCMD:
		Munsch.stMunschCmd.etCommand := ET_MUNSCH_CMD_SETAIRTEMP;
		Munsch.stMunschCmd.nAirTemp := nAirTemp;

		etMunschExtruder := ET_MunschExtruder_eExecuteCMD;              (* Next step *)

	ET_MunschExtruder_eExecuteCMD:
		nWatchdog := nWatchdog + 1;

		Munsch.bSendExe := TRUE;

		IF Munsch.bStringReceived
		THEN
			IF Munsch.stMunschRes.etResponse = ET_MUNSCH_RES_SETAIRTEMP
			     AND Munsch.stMunschCmd.nAirTemp = Munsch.stMunschRes.nAirRefTemp
			THEN
				Munsch.bSendExe := FALSE;

				nWatchdog := 0;

				etMunschExtruder := ET_MunschExtruder_eSetREQ;              (* Next step *)

			END_IF

		ELSIF Munsch.bInterfaceError
			    OR nWatchdog > 1000
		THEN
			Munsch.bSendExe := FALSE;

			udnErrorNo := 2;                     (* Error number *)
			etMunschExtruder := ET_MunschExtruder_eError;              (* Next step *)

		END_IF

	ET_MunschExtruder_eSetREQ:
		Munsch.stMunschCmd.etCommand := ET_MUNSCH_CMD_REQAIRREFTEMP;

		etMunschExtruder := ET_MunschExtruder_eExecuteREQ;              (* Next step *)

	ET_MunschExtruder_eExecuteREQ:
		nWatchdog := nWatchdog + 1;

		Munsch.bSendExe := TRUE;

		IF Munsch.bStringReceived
		THEN
			IF Munsch.stMunschRes.etResponse = ET_MUNSCH_RES_REQAIRREFTEMP
			THEN
				Munsch.nAirRefTemp := Munsch.stMunschRes.nAirRefTemp;

				Munsch.bSendExe := FALSE;

				nWatchdog := 0;
				etMunschExtruder := ET_MunschExtruder_eDone;              (* Next step *)
			END_IF

		ELSIF Munsch.bInterfaceError
			    OR nWatchdog > 1000
		THEN
			Munsch.bSendExe := FALSE;

			udnErrorNo := 3;                     (* Error number *)
			etMunschExtruder := ET_MunschExtruder_eError;              (* Next step *)

		END_IF

	ET_MunschExtruder_eError:
		bBusy := FALSE;						(* Command busy *)
		bError := TRUE;						(* Command error  *)

		etMunschExtruder := ET_MunschExtruder_eNoExecute;

	ET_MunschExtruder_eDone:
		bDone := TRUE;						(* Command done *)
		bBusy := FALSE;						(* Command busy *)

		etMunschExtruder := ET_MunschExtruder_eNoExecute;

	ET_MunschExtruder_eNoExecute:
		IF NOT bExecute
		THEN
			(* Reset outputs *)
			bDone := FALSE;						(* Command done *)
			bBusy := FALSE;						(* Command busy *)
			bError := FALSE;						(* Command error  *)

			nWatchdog := 0;
			Munsch.bLockedInterface := FALSE;

			Munsch.stMunschCmd.etCommand := ET_MUNSCH_CMD_NOCMD;
			Munsch.stMunschRes.etResponse := ET_MUNSCH_RES_NOCMD;

			etMunschExtruder := ET_MunschExtruder_eWaitExecute;
		END_IF
END_CASE;

bAirTempAlarm := Munsch.nAirActTemp > Munsch.nAirRefTemp + nAirTempTolerance
				OR Munsch.nAirActTemp > Munsch.nAirRefTemp - nAirTempTolerance;

END_FUNCTION_BLOCK

// ---- POUs/Tc3 Objects/ExternalHardware/Munsch/FB_MunschExtruder_Heat_1.TcPOU
FUNCTION_BLOCK FB_MunschExtruder_Heat_1
(*

The function block used to control heating Munsch extruder

Constructor: 		Patryk Panylo
Company:		E. Riexinger GmbH
Date:			13.10.2015
Version:			1.00

Date:			Revision:		Who:				Comment
dd.mm.yyyy		x.xx			Initials			comment

*)
VAR_INPUT
	(* Input variables / Eingang Variablen *)
	bEnable						:BOOL;						(* Enable FB signal *)
	bExtruderAirOk				:BOOL;						(* Signal extruder air ok *)
	bStart						:BOOL;						(* Start heating *)
	bStop						:BOOL;						(* Start heating *)
	nMaterialTemp				:INT;						(* Material temperatur *)
	nMinMaterialTemp			:INT;						(* Minimal material temperatur *)
	nMaxMaterialTemp			:INT;						(* Maximal material temperatur *)
	nAirTemp					:INT;						(* Air temperatur *)
	nMinAirTemp					:INT;						(* Minimal air temperatur *)
	nMaxAirTemp				:INT;						(* Maximal air temperatur *)
	tTimeOutAir					:TIME := t#30s;				(* Timeout of air ok *)
END_VAR
VAR_OUTPUT
	(* Output variables / Ausgang Variablen *)
	bExtruderAirOn				:BOOL;						(* Extruder air on*)
	bDone						:BOOL;						(* Program done *)
	bBusy						:BOOL;						(* Program busy *)
	bError						:BOOL;						(* Error *)
	udnErrorNo					:UDINT;
END_VAR
VAR_IN_OUT
	(* Input Output variables / Ausgang Variablen *)
	Munsch						:ST_MUNSCH_REF;
END_VAR
VAR
	(* Enummerations *)
	etMunschExtruder				:ET_MunschExtruder;

	(* Variables *)
	nWatchdog					:INT;

	(* References *)

	(* Interfaces *)

	(* Instances *)
	fbMaterialTemp				:FB_MunschExtruder_MaterialTemp;
	fbAirTemp					:FB_MunschExtruder_AirTemp;
	rtStart						:R_TRIG;
	rtStop						:R_TRIG;
	tonWatchdog					:TON;
END_VAR

IF NOT bEnable
THEN
	bDone := FALSE;					(* Program done *)
	bBusy := FALSE;                                  	(* Program not busy *)
	bError := FALSE;                                 	(* Program not error *)
	udnErrorNo := 0;                                 		(* Error number *)

	fbMaterialTemp(
		bEnable := FALSE,
		Munsch := Munsch
	);

	fbAirTemp(
		bEnable := FALSE,
		Munsch := Munsch
	);

	tonWatchdog(IN := FALSE);

	bExtruderAirOn := FALSE;
	Munsch.bHeat := FALSE;

	RETURN;
END_IF;

(* Wait for triger *)
rtStart(
	CLK := bStart
);

rtStop(
	CLK := bStop
);

IF  NOT Munsch.bHeat
THEN
	Munsch.nExtrudingSpeed := 0;
END_IF

IF rtStop.Q
THEN
	Munsch.bSetAirTemp := FALSE;
	Munsch.bSetMaterialTemp := FALSE;
	Munsch.bStartHeat := FALSE;
	Munsch.bStopHeat  := TRUE;
	Munsch.bStartExtruding := FALSE;
	Munsch.bStopExtruding  := FALSE;
	Munsch.bReadStatus := FALSE;

	Munsch.nExtrudingSpeed := 0;
END_IF

(* Send command *)
CASE etMunschExtruder OF

	ET_MunschExtruder_eWaitExecute:
		IF rtStop.Q
		    OR Munsch.bStopHeat
		THEN
			nWatchdog := 0;

			Munsch.bSetAirTemp := FALSE;
			Munsch.bSetMaterialTemp := FALSE;
			Munsch.bStartHeat := FALSE;
			Munsch.bStopHeat  := TRUE;
			Munsch.bStartExtruding := FALSE;
			Munsch.bStopExtruding  := FALSE;
			Munsch.bReadStatus := FALSE;

			Munsch.nExtrudingSpeed := 0;

			etMunschExtruder := ET_MunschExtruder_eChkInterface;              (* Next step *)

		ELSIF rtStart.Q
		THEN
			nWatchdog := 0;

			Munsch.bSetAirTemp := FALSE;
			Munsch.bSetMaterialTemp := FALSE;
			Munsch.bStartHeat := TRUE;
			Munsch.bStopHeat  := FALSE;
			Munsch.bStartExtruding := FALSE;
			Munsch.bStopExtruding  := FALSE;
			Munsch.bReadStatus := FALSE;

			etMunschExtruder := ET_MunschExtruder_eChkInterface;              (* Next step *)

		END_IF

	ET_MunschExtruder_eChkInterface:
		nWatchdog := nWatchdog + 1;

		IF NOT Munsch.bLockedInterface
		THEN
			bBusy := FALSE;                                     	(* Program not busy *)
			bError := FALSE;                         		(* Program not error *)
			udnErrorNo := 0;                         		(* Error number *)

			IF Munsch.bStopHeat
			THEN
				nWatchdog := 0;
				bDone:= FALSE;                               		(* Program done *)
				bBusy := TRUE;                                  	(* Program busy *)
	
				bExtruderAirOn := FALSE;
				tonWatchdog(IN := FALSE);
	
				Munsch.bLockedInterface := TRUE;
				Munsch.bSendExe := FALSE;
	
				etMunschExtruder := ET_MunschExtruder_eSetCMD;              (* Next step *)
	
			ELSIF Munsch.bStartHeat
			THEN
				nWatchdog := 0;
				bDone:= FALSE;                               		(* Program done *)
				bBusy := TRUE;                                  	(* Program busy *)
	
				fbMaterialTemp(
					bEnable := TRUE,
					bExecute := FALSE,
					nMaterialTemp := nMaterialTemp,
					nMinMaterialTemp := nMinMaterialTemp,
					nMaxMaterialTemp := nMaxMaterialTemp,
					Munsch := Munsch
				);
				
				fbAirTemp(
					bEnable := TRUE,
					bExecute := FALSE,
					nAirTemp := nAirTemp,
					nMinAirTemp := nMinAirTemp,
					nMaxAirTemp := nMaxAirTemp,
					Munsch := Munsch
				);
	
				bExtruderAirOn := TRUE;
				tonWatchdog(IN := FALSE);

				Munsch.bLockedInterface := TRUE;
				Munsch.bSendExe := FALSE;

				etMunschExtruder := ET_MunschExtruder_eSetCMD;              (* Next step *)

			ELSE
				etMunschExtruder :=  ET_MunschExtruder_eError;             (* Next step *)
			END_IF

			Munsch.bStartHeat := FALSE;
			Munsch.bStopHeat  := FALSE;

		ELSIF nWatchdog > 1000
		THEN
			Munsch.bStartHeat := FALSE;
			Munsch.bStopHeat  := FALSE;

